DATA_BLOCK "DB_ALARM"   // DB100
{ S7_Optimized_Access := 'FALSE' }
// stored: AutoNumber false
   VAR
      ALARM : Struct
         ALARM_GLOBAL : Bool;   // globální alarm
         HERMA_ERROR : Bool;
         ALARM_2 : Bool;
         ALARM_3 : Bool;
         ALARM_4 : Bool;
         ALARM_5 : Bool;
         air : Bool;   // nedostatečný tlak vzduchu
         ALARM_7 : Bool;
         ALARM_8 : Bool;
         ALARM_9 : Bool;
         ALARM_10 : Bool;
         ALARM_11 : Bool;
         ALARM_12 : Bool;
         ALARM_13 : Bool;
         ALARM_14 : Bool;
         vypadek_safety_karty : Bool;
      END_STRUCT;
      WRONG : Struct
         NENI_INICIALIZACE : Bool;
         WRONG_global : Bool;
         dvere_L_tevreny : Bool;
         dvere_P_otevreny : Bool;
         WRONG_4 : Bool;
         WRONG_5 : Bool;
         WRONG_6 : Bool;
         WRONG_7 : Bool;
         WRONG_8 : Bool;
         WRONG_9 : Bool;
         WRONG_10 : Bool;
         WRONG_11 : Bool;
         WRONG_12 : Bool;
         WRONG_13 : Bool;
         rop_glob_warning : Bool;
         rop_active_autocale : Bool;
      END_STRUCT;
      OP0 : Struct
         ALARM : Struct
            DOOR_ERROR : Bool;
            ALARM_1 : Bool;
            ALARM_2 : Bool;
            ALARM_3 : Bool;
            ALARM_4 : Bool;
            ALARM_5 : Bool;
            ALARM_6 : Bool;
            ALARM_7 : Bool;
            ALARM_8 : Bool;
            ALARM_9 : Bool;
            ALARM_10 : Bool;
            ALARM_11 : Bool;
            ALARM_12 : Bool;
            ALARM_13 : Bool;
            ALARM_14 : Bool;
            ALARM_15 : Bool;
         END_STRUCT;
         WRONG : Struct
            WRONG_0 : Bool;
            WRONG_1 : Bool;
            WRONG_2 : Bool;
            WRONG_3 : Bool;
            WRONG_4 : Bool;
            WRONG_5 : Bool;
            WRONG_6 : Bool;
            WRONG_7 : Bool;
            WRONG_8 : Bool;
            WRONG_9 : Bool;
            WRONG_10 : Bool;
            WRONG_11 : Bool;
            WRONG_12 : Bool;
            WRONG_13 : Bool;
            WRONG_14 : Bool;
            WRONG_15 : Bool;
         END_STRUCT;
         M_0 : Int;
         M_1 : Int;
         M_2 : Int;
         M_3 : Int;
         M_4 : Int;
         M_5 : Int;
         M_6 : Int;
         M_7 : Int;
         M_8 : Int;
         M_9 : Int;
         M_10 : Int;
         M_11 : Int;
         M_12 : Int;
         M_13 : Int;
         M_14 : Int;
         M_15 : Int;
      END_STRUCT;
      OP1 : Struct
         ALARM : Struct
            dvere_1 : Bool;
            ALARM_1 : Bool;
            ALARM_2 : Bool;
            ALARM_3 : Bool;
            ALARM_4 : Bool;
            ALARM_5 : Bool;
            ALARM_6 : Bool;
            hladina_mimo_mez : Bool;
            ALARM_8 : Bool;
            ALARM_9 : Bool;
            ALARM_10 : Bool;
            ALARM_11 : Bool;
            ALARM_12 : Bool;
            ALARM_13 : Bool;
            ALARM_14 : Bool;
            ALARM_15 : Bool;
         END_STRUCT;
         WRONG : Struct
            WRONG_0 : Bool;
            WRONG_1 : Bool;
            WRONG_2 : Bool;
            WRONG_3 : Bool;
            WRONG_4 : Bool;
            WRONG_5 : Bool;
            WRONG_6 : Bool;
            WRONG_7 : Bool;
            WRONG_8 : Bool;
            WRONG_9 : Bool;
            WRONG_10 : Bool;
            WRONG_11 : Bool;
            WRONG_12 : Bool;
            WRONG_13 : Bool;
            WRONG_14 : Bool;
            WRONG_15 : Bool;
         END_STRUCT;
         "-Y7_KARUSEL" : Int;
         "-Y9_ZARAZKA" : Int;
         M_2 : Int;
         M_3 : Int;
         M_4 : Int;
         M_5 : Int;
         M_6 : Int;
         M_7 : Int;
         M_8 : Int;
         M_9 : Int;
         M_10 : Int;
         M_11 : Int;
         M_12 : Int;
         M_13 : Int;
         M_14 : Int;
         M_15 : Int;
      END_STRUCT;
      OP2 : Struct
         ALARM : Struct
            dvere_1 : Bool;
            dvere_2 : Bool;
            dvere_3 : Bool;
            dvere_4 : Bool;
            paprsek : Bool;
            porucha_svarovani : Bool;
            rop_alarm : Bool;
            servo_power_error : Bool;
            servo_jog_error : Bool;
            servo_homing : Bool;
            Cel_podel_porucha : Bool;
            vysoka_tuzka : Bool;
            ALARM_12 : Bool;
            ALARM_13 : Bool;
            folie : Bool;
            ALARM_15 : Bool;
         END_STRUCT;
         WRONG : Struct
            WRONG_0 : Bool;
            WRONG_1 : Bool;
            WRONG_2 : Bool;
            WRONG_3 : Bool;
            WRONG_4 : Bool;
            WRONG_5 : Bool;
            WRONG_6 : Bool;
            WRONG_7 : Bool;
            WRONG_8 : Bool;
            WRONG_9 : Bool;
            WRONG_10 : Bool;
            WRONG_11 : Bool;
            WRONG_12 : Bool;
            WRONG_13 : Bool;
            WRONG_14 : Bool;
            WRONG_15 : Bool;
         END_STRUCT;
         A1 : Int;   // -YA1
         A2 : Int;   // -YA2
         A3 : Int;   // -YA3
         A4 : Int;   // -YA4
         A5 : Int;   // -YA5
         A6 : Int;   // -YA6
         A7 : Int;   // -YA7
         A8 : Int;   // -YA8
         M_8 : Int;
         M_9 : Int;
         M_10 : Int;
         M_11 : Int;
         M_12 : Int;
         M_13 : Int;
         M_14 : Int;
         M_15 : Int;
      END_STRUCT;
      OP3 : Struct
         ALARM : Struct
            ALARM_0 : Bool;
            ALARM_1 : Bool;
            ALARM_2 : Bool;
            ALARM_3 : Bool;
            ALARM_4 : Bool;
            ALARM_5 : Bool;
            ALARM_6 : Bool;
            ALARM_7 : Bool;
            ALARM_8 : Bool;
            ALARM_9 : Bool;
            ALARM_10 : Bool;
            ALARM_11 : Bool;
            ALARM_12 : Bool;
            ALARM_13 : Bool;
            ALARM_14 : Bool;
            ALARM_15 : Bool;
         END_STRUCT;
         WRONG : Struct
            WRONG_0 : Bool;
            WRONG_1 : Bool;
            WRONG_2 : Bool;
            WRONG_3 : Bool;
            WRONG_4 : Bool;
            WRONG_5 : Bool;
            WRONG_6 : Bool;
            WRONG_7 : Bool;
            WRONG_8 : Bool;
            WRONG_9 : Bool;
            WRONG_10 : Bool;
            WRONG_11 : Bool;
            WRONG_12 : Bool;
            WRONG_13 : Bool;
            WRONG_14 : Bool;
            WRONG_15 : Bool;
         END_STRUCT;
         B1 : Int;   // -YB1
         B2 : Int;   // -YB2
         B3 : Int;   // -YB3
         B4 : Int;   // -YB4
         B5 : Int;   // -YB5
         B6 : Int;   // -YB6
         B7 : Int;   // -YB7
         B8 : Int;   // -YB8
         M_8 : Int;
         M_9 : Int;
         M_10 : Int;
         M_11 : Int;
         M_12 : Int;
         M_13 : Int;
         M_14 : Int;
         M_15 : Int;
      END_STRUCT;
      OP4 : Struct
         ALARM : Struct
            odsavani_nefunguje : Bool;
            ALARM_1 : Bool;
            ALARM_2 : Bool;
            ALARM_3 : Bool;
            ALARM_4 : Bool;
            ALARM_5 : Bool;
            ALARM_6 : Bool;
            ALARM_7 : Bool;
            ALARM_8 : Bool;
            ALARM_9 : Bool;
            ALARM_10 : Bool;
            ALARM_11 : Bool;
            ALARM_12 : Bool;
            ALARM_13 : Bool;
            ALARM_14 : Bool;
            ALARM_15 : Bool;
         END_STRUCT;
         WRONG : Struct
            WRONG_0 : Bool;
            WRONG_1 : Bool;
            WRONG_2 : Bool;
            WRONG_3 : Bool;
            WRONG_4 : Bool;
            WRONG_5 : Bool;
            WRONG_6 : Bool;
            WRONG_7 : Bool;
            WRONG_8 : Bool;
            WRONG_9 : Bool;
            WRONG_10 : Bool;
            WRONG_11 : Bool;
            WRONG_12 : Bool;
            WRONG_13 : Bool;
            WRONG_14 : Bool;
            WRONG_15 : Bool;
         END_STRUCT;
         M_0 : Int;
         M_1 : Int;
         M_2 : Int;
         M_3 : Int;
         M_4 : Int;
         M_5 : Int;
         M_6 : Int;
         M_7 : Int;
         M_8 : Int;
         M_9 : Int;
         M_10 : Int;
         M_11 : Int;
         M_12 : Int;
         M_13 : Int;
         M_14 : Int;
         M_15 : Int;
      END_STRUCT;
      OP5 : Struct
         ALARM : Struct
            ALARM_0 : Bool;
            ALARM_1 : Bool;
            ALARM_2 : Bool;
            ALARM_3 : Bool;
            ALARM_4 : Bool;
            ALARM_5 : Bool;
            ALARM_6 : Bool;
            ALARM_7 : Bool;
            ALARM_8 : Bool;
            ALARM_9 : Bool;
            ALARM_10 : Bool;
            ALARM_11 : Bool;
            ALARM_12 : Bool;
            ALARM_13 : Bool;
            ALARM_14 : Bool;
            ALARM_15 : Bool;
         END_STRUCT;
         WRONG : Struct
            WRONG_0 : Bool;
            WRONG_1 : Bool;
            WRONG_2 : Bool;
            WRONG_3 : Bool;
            WRONG_4 : Bool;
            WRONG_5 : Bool;
            WRONG_6 : Bool;
            WRONG_7 : Bool;
            WRONG_8 : Bool;
            WRONG_9 : Bool;
            WRONG_10 : Bool;
            WRONG_11 : Bool;
            WRONG_12 : Bool;
            WRONG_13 : Bool;
            WRONG_14 : Bool;
            WRONG_15 : Bool;
         END_STRUCT;
         M_0 : Int;
         M_1 : Int;
         M_2 : Int;
         M_3 : Int;
         M_4 : Int;
         M_5 : Int;
         M_6 : Int;
         M_7 : Int;
         M_8 : Int;
         M_9 : Int;
         M_10 : Int;
         M_11 : Int;
         M_12 : Int;
         M_13 : Int;
         M_14 : Int;
         M_15 : Int;
      END_STRUCT;
      null : Struct
         ALARM_0 : Bool;
         ALARM_1 : Bool;
         ALARM_2 : Bool;
         ALARM_3 : Bool;
         ALARM_4 : Bool;
         ALARM_5 : Bool;
         ALARM_6 : Bool;
         ALARM_7 : Bool;
         ALARM_8 : Bool;
         ALARM_9 : Bool;
         ALARM_10 : Bool;
         ALARM_11 : Bool;
         ALARM_12 : Bool;
         ALARM_13 : Bool;
         ALARM_14 : Bool;
         ALARM_15 : Bool;
      END_STRUCT;
      alarmy : Array[0..255] of Bool;
      alarm_line : Int;
      wrong_line : Int;
      alarm_op_1 : Int;
      wrong_op_1 : Int;
      alarm_op_2 : Int;
      wrong_op_2 : Int;
      alarm_op_3 : Int;
      wrong_op_3 : Int;
      alarm_op_4 : Int;
      wrong_op_4 : Int;
      alarm_op_5 : Int;
      wrong_op_5 : Int;
      T_tiskarna : TON_TIME;
   END_VAR
BEGIN
END_DATA_BLOCK

DATA_BLOCK "DB_STS_M"   // DB101
{ S7_Optimized_Access := 'FALSE' }
// stored: AutoNumber false
   VAR
      OP0 : Struct
         STS_M0 : UInt;
         STS_M1 : UInt;
         STS_M2 : UInt;
         STS_M3 : UInt;
         STS_M4 : UInt;
         STS_M5 : UInt;
         STS_M6 : UInt;
         STS_M7 : UInt;
         STS_M8 : UInt;
         STS_M9 : UInt;
         STS_M10 : UInt;
         STS_M11 : UInt;
         STS_M12 : UInt;
         STS_M13 : UInt;
         STS_M14 : UInt;
         STS_M15 : UInt;
      END_STRUCT;
      OP1 : Struct
         KARUSEL : UInt;
         ZARAZKA : UInt;
         STS_M2 : UInt;
         STS_M3 : UInt;
         STS_M4 : UInt;
         STS_M5 : UInt;
         STS_M6 : UInt;
         STS_M7 : UInt;
         STS_M8 : UInt;
         STS_M9 : UInt;
         STS_M10 : UInt;
         STS_M11 : UInt;
         STS_M12 : UInt;
         STS_M13 : UInt;
         STS_M14 : UInt;
         STS_M15 : UInt;
         OP1 : Struct
            STS_M0 : UInt;
            STS_M1 : UInt;
            STS_M2 : UInt;
            STS_M3 : UInt;
            STS_M4 : UInt;
            STS_M5 : UInt;
            STS_M6 : UInt;
            STS_M7 : UInt;
            STS_M8 : UInt;
            STS_M9 : UInt;
            STS_M10 : UInt;
            STS_M11 : UInt;
            STS_M12 : UInt;
            STS_M13 : UInt;
            STS_M14 : UInt;
            STS_M15 : UInt;
         END_STRUCT;
      END_STRUCT;
      OP2 : Struct
         A1 : UInt;
         A2 : UInt;
         A3 : UInt;
         A4 : UInt;
         A5 : UInt;
         A6 : UInt;
         A7 : UInt;
         A8 : UInt;
         STS_M8 : UInt;
         STS_M9 : UInt;
         STS_M10 : UInt;
         STS_M11 : UInt;
         STS_M12 : UInt;
         STS_M13 : UInt;
         STS_M14 : UInt;
         STS_M15 : UInt;
      END_STRUCT;
      OP3 : Struct
         B1 : UInt;
         B2 : UInt;
         B3 : UInt;
         B4 : UInt;
         B5 : UInt;
         B6 : UInt;
         B7 : UInt;
         B8 : UInt;
         STS_M8 : UInt;
         STS_M9 : UInt;
         STS_M10 : UInt;
         STS_M11 : UInt;
         STS_M12 : UInt;
         STS_M13 : UInt;
         STS_M14 : UInt;
         STS_M15 : UInt;
      END_STRUCT;
   END_VAR
BEGIN
END_DATA_BLOCK

DATA_BLOCK "DB_DATA_LASER"   // DB401
{ S7_Optimized_Access := 'TRUE' }
// stored: AutoNumber false, MemoryReserve 100
   VAR
      LASER_DATA_READ : Array[0..71] of Byte;
      LASER_DATA_WRITE : Array[0..71] of Byte;
      READ : Bool;
      WRITE : Bool;
   END_VAR
BEGIN
END_DATA_BLOCK

DATA_BLOCK "DB_LASER"   // DB402
{ S7_Optimized_Access := 'TRUE' }
// stored: AutoNumber false, MemoryReserve 100
   VAR
      DATA_DO_ETIKETY : Struct
         TEXT : String[5];
         "INT" : Int;
         "REAL" : Real;
         PROGRAM : Array[0..1] of String[10];
      END_STRUCT;
      DATA_DO_DAT : Struct
         ZAVORKA_L : Char := '<';
         ZAVORKA_P : Char := '>';
         XLP : Array[0..3] of Char;
      END_STRUCT;
      smaz_me_start : Bool;
      smaz_me_adresa : Int;
   END_VAR
BEGIN
   DATA_DO_ETIKETY.PROGRAM[0] := 'TEST_1';
   DATA_DO_ETIKETY.PROGRAM[1] := 'TEST_222';
   DATA_DO_DAT.XLP[0] := '.';
   DATA_DO_DAT.XLP[1] := 'x';
   DATA_DO_DAT.XLP[2] := 'l';
   DATA_DO_DAT.XLP[3] := 'p';
END_DATA_BLOCK

ORGANIZATION_BLOCK "Main"   // OB1, LAD, ProgramCycle
TITLE = "Main Program Sweep (Cycle)"
{ S7_Optimized_Access := 'TRUE' }
// stored: SetENOAutomatically false
   VAR_INPUT
      Initial_Call : Bool;   // Initial call of this OB
      Remanence : Bool;   // =True, if remanent data are available
   END_VAR
BEGIN

REGION Network 1
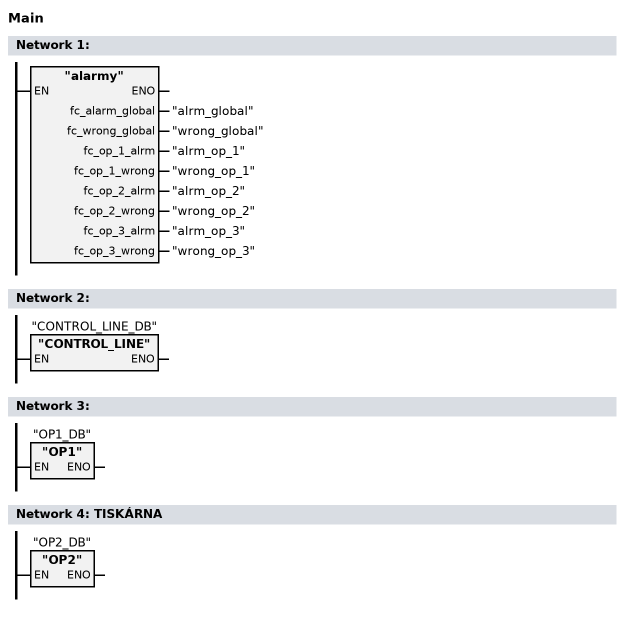
   RUNG wire#powerrail
      "alarmy"(fc_alarm_global => "alrm_global", fc_wrong_global => "wrong_global", fc_op_1_alrm => "alrm_op_1", fc_op_1_wrong => "wrong_op_1", fc_op_2_alrm => "alrm_op_2", fc_op_2_wrong => "wrong_op_2", fc_op_3_alrm => "alrm_op_3", fc_op_3_wrong => "wrong_op_3")
   END_RUNG
   // the same network as SCL:
   "alarmy"(fc_alarm_global => "alrm_global",
            fc_wrong_global => "wrong_global",
            fc_op_1_alrm => "alrm_op_1",
            fc_op_1_wrong => "wrong_op_1",
            fc_op_2_alrm => "alrm_op_2",
            fc_op_2_wrong => "wrong_op_2",
            fc_op_3_alrm => "alrm_op_3",
            fc_op_3_wrong => "wrong_op_3");
END_REGION

REGION Network 2
   RUNG wire#powerrail
      "CONTROL_LINE_DB"()
   END_RUNG
   // the same network as SCL:
   "CONTROL_LINE_DB"();   // "CONTROL_LINE"
END_REGION

REGION Network 3
   RUNG wire#powerrail
      "OP1_DB"()
   END_RUNG
   // the same network as SCL:
   "OP1_DB"();   // "OP1"
END_REGION

REGION Network 4: TISKÁRNA
   RUNG wire#powerrail
      "OP2_DB"()
   END_RUNG
   // the same network as SCL:
   "OP2_DB"();   // "OP2"
END_REGION
END_ORGANIZATION_BLOCK

FUNCTION "alarmy" : Void   // FC100, LAD
{ S7_Optimized_Access := 'TRUE' }
// stored: AutoNumber false, SetENOAutomatically false
   VAR_OUTPUT
      fc_alarm_global : Bool;
      fc_wrong_global : Bool;
      fc_op_1_alrm : Bool;
      fc_op_1_wrong : Bool;
      fc_op_2_alrm : Bool;
      fc_op_2_wrong : Bool;
      fc_op_3_alrm : Bool;
      fc_op_3_wrong : Bool;
   END_VAR
   VAR_TEMP
      OP_1_E : Bool;
      OP_2_E : Bool;
      OP_3_E : Bool;
      OP_4_E : Bool;
      OP_5_E : Bool;
      OP_1_W : Bool;
      OP_2_W : Bool;
      OP_3_W : Bool;
      OP_4_W : Bool;
      OP_5_W : Bool;
   END_VAR
   VAR CONSTANT
      TIME_ERROR_BOR : Time := T#4S;
   END_VAR
BEGIN

REGION Network 1: op_1 alarmy proces
END_REGION

REGION Network 2: op_1_warning_proces
END_REGION

REGION Network 3: OP_1_ALARM
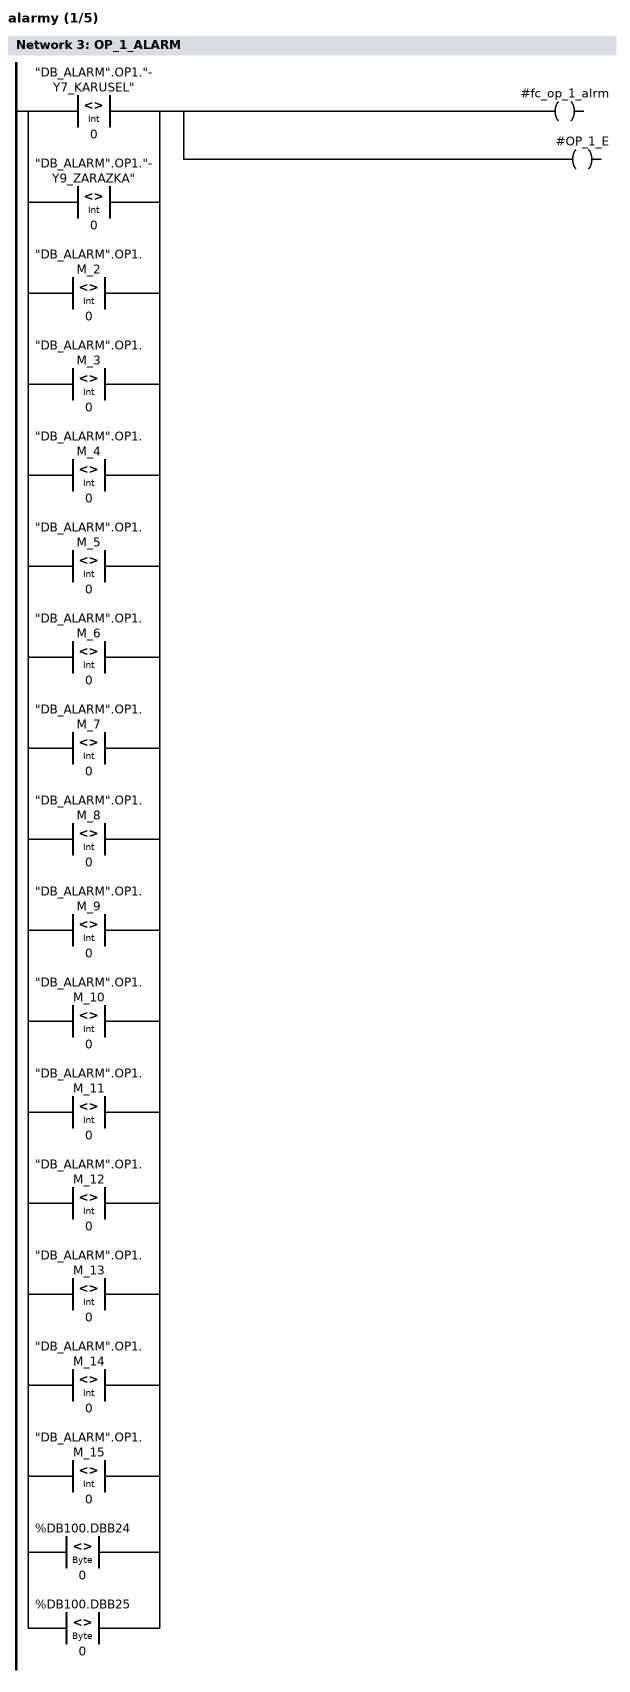
   RUNG wire#powerrail
      { S7_Templates := "SrcType := Int" } NE_Contact(in1 := "DB_ALARM".OP1."-Y7_KARUSEL", in2 := 0)
      wire#w1
      Coil( #fc_op_1_alrm )
   END_RUNG
   RUNG wire#powerrail
      { S7_Templates := "SrcType := Int" } NE_Contact(in1 := "DB_ALARM".OP1."-Y9_ZARAZKA", in2 := 0)
   END_RUNG wire#w1
   RUNG wire#powerrail
      { S7_Templates := "SrcType := Int" } NE_Contact(in1 := "DB_ALARM".OP1.M_2, in2 := 0)
   END_RUNG wire#w1
   RUNG wire#powerrail
      { S7_Templates := "SrcType := Int" } NE_Contact(in1 := "DB_ALARM".OP1.M_3, in2 := 0)
   END_RUNG wire#w1
   RUNG wire#powerrail
      { S7_Templates := "SrcType := Int" } NE_Contact(in1 := "DB_ALARM".OP1.M_4, in2 := 0)
   END_RUNG wire#w1
   RUNG wire#powerrail
      { S7_Templates := "SrcType := Int" } NE_Contact(in1 := "DB_ALARM".OP1.M_5, in2 := 0)
   END_RUNG wire#w1
   RUNG wire#powerrail
      { S7_Templates := "SrcType := Int" } NE_Contact(in1 := "DB_ALARM".OP1.M_6, in2 := 0)
   END_RUNG wire#w1
   RUNG wire#powerrail
      { S7_Templates := "SrcType := Int" } NE_Contact(in1 := "DB_ALARM".OP1.M_7, in2 := 0)
   END_RUNG wire#w1
   RUNG wire#powerrail
      { S7_Templates := "SrcType := Int" } NE_Contact(in1 := "DB_ALARM".OP1.M_8, in2 := 0)
   END_RUNG wire#w1
   RUNG wire#powerrail
      { S7_Templates := "SrcType := Int" } NE_Contact(in1 := "DB_ALARM".OP1.M_9, in2 := 0)
   END_RUNG wire#w1
   RUNG wire#powerrail
      { S7_Templates := "SrcType := Int" } NE_Contact(in1 := "DB_ALARM".OP1.M_10, in2 := 0)
   END_RUNG wire#w1
   RUNG wire#powerrail
      { S7_Templates := "SrcType := Int" } NE_Contact(in1 := "DB_ALARM".OP1.M_11, in2 := 0)
   END_RUNG wire#w1
   RUNG wire#powerrail
      { S7_Templates := "SrcType := Int" } NE_Contact(in1 := "DB_ALARM".OP1.M_12, in2 := 0)
   END_RUNG wire#w1
   RUNG wire#powerrail
      { S7_Templates := "SrcType := Int" } NE_Contact(in1 := "DB_ALARM".OP1.M_13, in2 := 0)
   END_RUNG wire#w1
   RUNG wire#powerrail
      { S7_Templates := "SrcType := Int" } NE_Contact(in1 := "DB_ALARM".OP1.M_14, in2 := 0)
   END_RUNG wire#w1
   RUNG wire#powerrail
      { S7_Templates := "SrcType := Int" } NE_Contact(in1 := "DB_ALARM".OP1.M_15, in2 := 0)
   END_RUNG wire#w1
   RUNG wire#powerrail
      { S7_Templates := "SrcType := Byte" } NE_Contact(in1 := %DB100.DBB24, in2 := 0)
   END_RUNG wire#w1
   RUNG wire#powerrail
      { S7_Templates := "SrcType := Byte" } NE_Contact(in1 := %DB100.DBB25, in2 := 0)
   END_RUNG wire#w1
   RUNG wire#w1
      Coil( #OP_1_E )
   END_RUNG
   // the same network as SCL:
   #fc_op_1_alrm := ("DB_ALARM".OP1."-Y7_KARUSEL" <> 0) OR ("DB_ALARM".OP1."-Y9_ZARAZKA" <> 0) OR ("DB_ALARM".OP1.M_2 <> 0) OR ("DB_ALARM".OP1.M_3 <> 0) OR ("DB_ALARM".OP1.M_4 <> 0) OR ("DB_ALARM".OP1.M_5 <> 0) OR ("DB_ALARM".OP1.M_6 <> 0) OR ("DB_ALARM".OP1.M_7 <> 0) OR ("DB_ALARM".OP1.M_8 <> 0) OR ("DB_ALARM".OP1.M_9 <> 0) OR ("DB_ALARM".OP1.M_10 <> 0) OR ("DB_ALARM".OP1.M_11 <> 0) OR ("DB_ALARM".OP1.M_12 <> 0) OR ("DB_ALARM".OP1.M_13 <> 0) OR ("DB_ALARM".OP1.M_14 <> 0) OR ("DB_ALARM".OP1.M_15 <> 0) OR (%DB100.DBB24 <> 0) OR (%DB100.DBB25 <> 0);
   #OP_1_E := #fc_op_1_alrm;
END_REGION

REGION Network 4: OP_2_ALARM
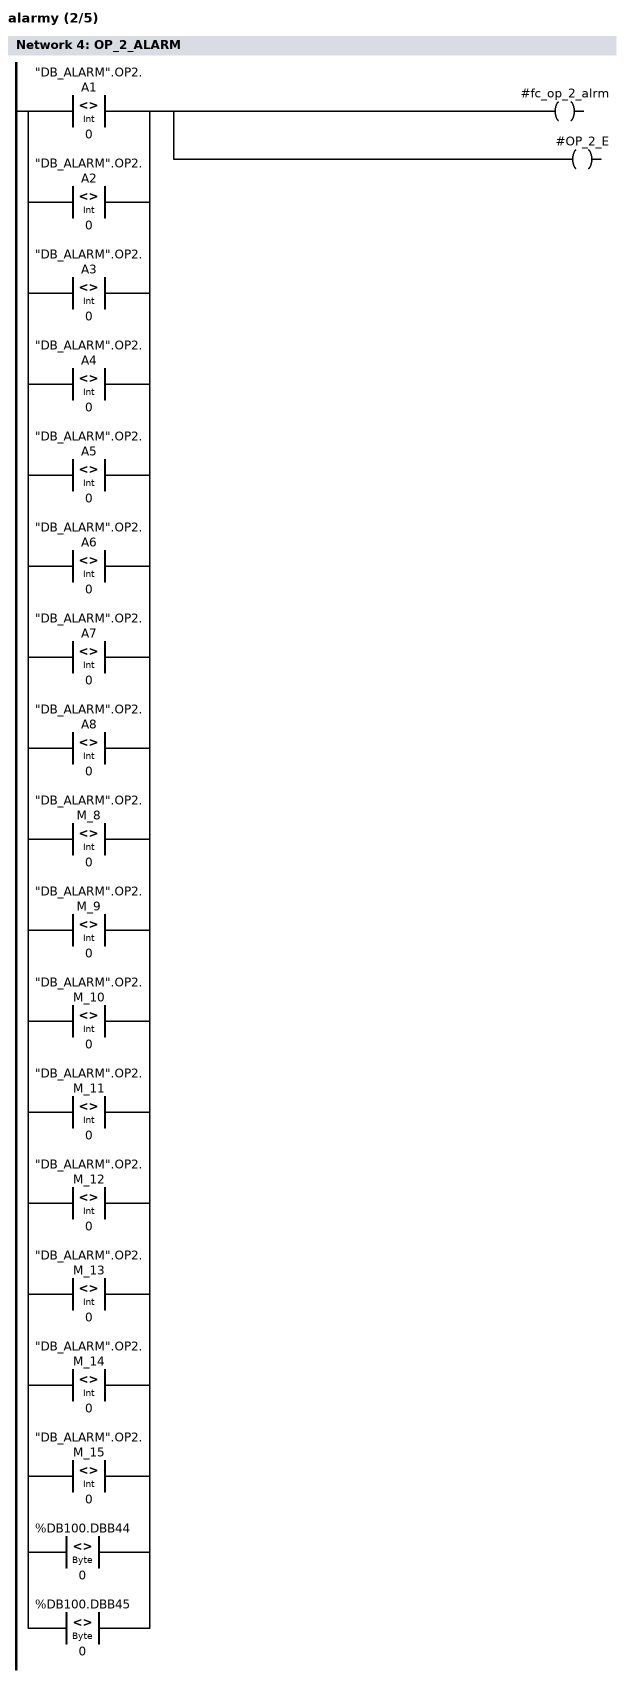
   RUNG wire#powerrail
      { S7_Templates := "SrcType := Int" } NE_Contact(in1 := "DB_ALARM".OP2.A1, in2 := 0)
      wire#w1
      Coil( #fc_op_2_alrm )
   END_RUNG
   RUNG wire#powerrail
      { S7_Templates := "SrcType := Int" } NE_Contact(in1 := "DB_ALARM".OP2.A2, in2 := 0)
   END_RUNG wire#w1
   RUNG wire#powerrail
      { S7_Templates := "SrcType := Int" } NE_Contact(in1 := "DB_ALARM".OP2.A3, in2 := 0)
   END_RUNG wire#w1
   RUNG wire#powerrail
      { S7_Templates := "SrcType := Int" } NE_Contact(in1 := "DB_ALARM".OP2.A4, in2 := 0)
   END_RUNG wire#w1
   RUNG wire#powerrail
      { S7_Templates := "SrcType := Int" } NE_Contact(in1 := "DB_ALARM".OP2.A5, in2 := 0)
   END_RUNG wire#w1
   RUNG wire#powerrail
      { S7_Templates := "SrcType := Int" } NE_Contact(in1 := "DB_ALARM".OP2.A6, in2 := 0)
   END_RUNG wire#w1
   RUNG wire#powerrail
      { S7_Templates := "SrcType := Int" } NE_Contact(in1 := "DB_ALARM".OP2.A7, in2 := 0)
   END_RUNG wire#w1
   RUNG wire#powerrail
      { S7_Templates := "SrcType := Int" } NE_Contact(in1 := "DB_ALARM".OP2.A8, in2 := 0)
   END_RUNG wire#w1
   RUNG wire#powerrail
      { S7_Templates := "SrcType := Int" } NE_Contact(in1 := "DB_ALARM".OP2.M_8, in2 := 0)
   END_RUNG wire#w1
   RUNG wire#powerrail
      { S7_Templates := "SrcType := Int" } NE_Contact(in1 := "DB_ALARM".OP2.M_9, in2 := 0)
   END_RUNG wire#w1
   RUNG wire#powerrail
      { S7_Templates := "SrcType := Int" } NE_Contact(in1 := "DB_ALARM".OP2.M_10, in2 := 0)
   END_RUNG wire#w1
   RUNG wire#powerrail
      { S7_Templates := "SrcType := Int" } NE_Contact(in1 := "DB_ALARM".OP2.M_11, in2 := 0)
   END_RUNG wire#w1
   RUNG wire#powerrail
      { S7_Templates := "SrcType := Int" } NE_Contact(in1 := "DB_ALARM".OP2.M_12, in2 := 0)
   END_RUNG wire#w1
   RUNG wire#powerrail
      { S7_Templates := "SrcType := Int" } NE_Contact(in1 := "DB_ALARM".OP2.M_13, in2 := 0)
   END_RUNG wire#w1
   RUNG wire#powerrail
      { S7_Templates := "SrcType := Int" } NE_Contact(in1 := "DB_ALARM".OP2.M_14, in2 := 0)
   END_RUNG wire#w1
   RUNG wire#powerrail
      { S7_Templates := "SrcType := Int" } NE_Contact(in1 := "DB_ALARM".OP2.M_15, in2 := 0)
   END_RUNG wire#w1
   RUNG wire#powerrail
      { S7_Templates := "SrcType := Byte" } NE_Contact(in1 := %DB100.DBB44, in2 := 0)
   END_RUNG wire#w1
   RUNG wire#powerrail
      { S7_Templates := "SrcType := Byte" } NE_Contact(in1 := %DB100.DBB45, in2 := 0)
   END_RUNG wire#w1
   RUNG wire#w1
      Coil( #OP_2_E )
   END_RUNG
   // the same network as SCL:
   #fc_op_2_alrm := ("DB_ALARM".OP2.A1 <> 0) OR ("DB_ALARM".OP2.A2 <> 0) OR ("DB_ALARM".OP2.A3 <> 0) OR ("DB_ALARM".OP2.A4 <> 0) OR ("DB_ALARM".OP2.A5 <> 0) OR ("DB_ALARM".OP2.A6 <> 0) OR ("DB_ALARM".OP2.A7 <> 0) OR ("DB_ALARM".OP2.A8 <> 0) OR ("DB_ALARM".OP2.M_8 <> 0) OR ("DB_ALARM".OP2.M_9 <> 0) OR ("DB_ALARM".OP2.M_10 <> 0) OR ("DB_ALARM".OP2.M_11 <> 0) OR ("DB_ALARM".OP2.M_12 <> 0) OR ("DB_ALARM".OP2.M_13 <> 0) OR ("DB_ALARM".OP2.M_14 <> 0) OR ("DB_ALARM".OP2.M_15 <> 0) OR (%DB100.DBB44 <> 0) OR (%DB100.DBB45 <> 0);
   #OP_2_E := #fc_op_2_alrm;
END_REGION

REGION Network 5: OP_3_ALARM
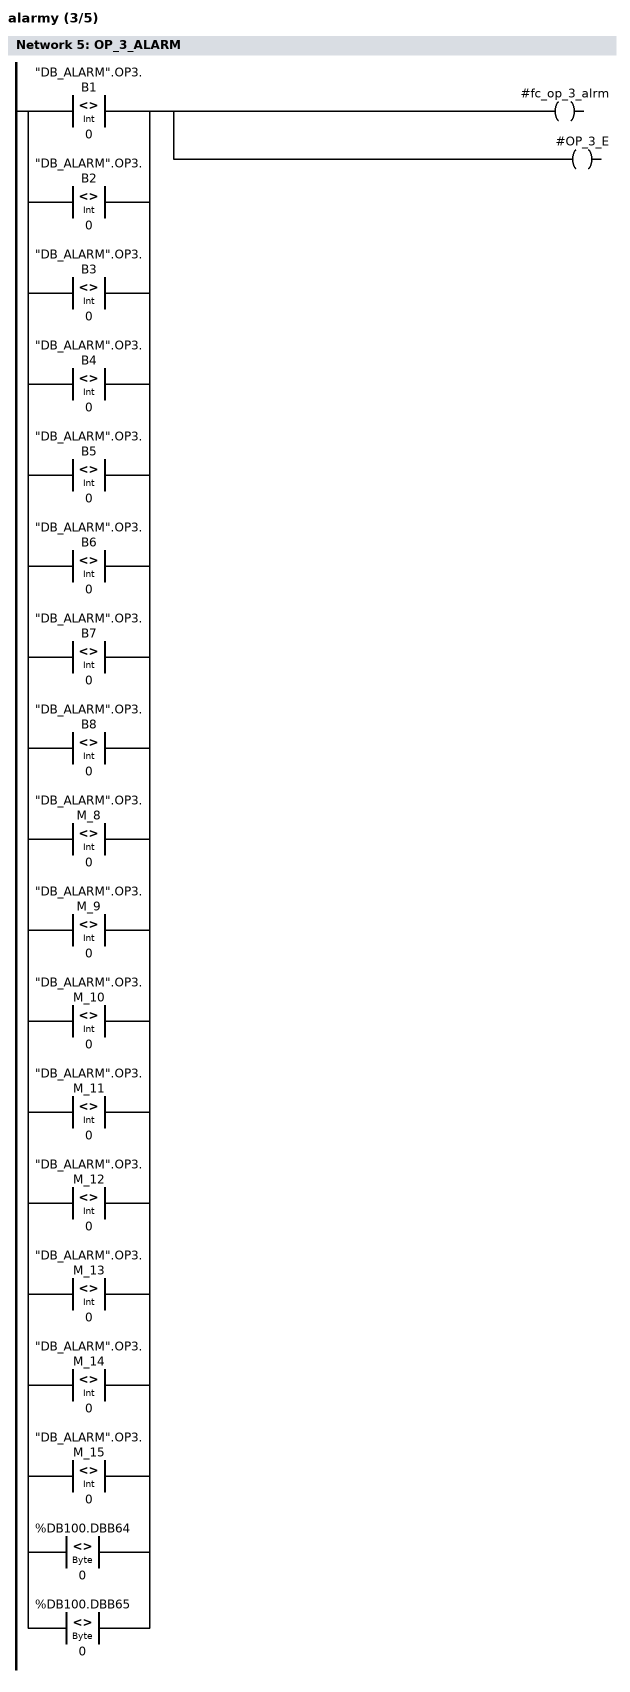
   RUNG wire#powerrail
      { S7_Templates := "SrcType := Int" } NE_Contact(in1 := "DB_ALARM".OP3.B1, in2 := 0)
      wire#w1
      Coil( #fc_op_3_alrm )
   END_RUNG
   RUNG wire#powerrail
      { S7_Templates := "SrcType := Int" } NE_Contact(in1 := "DB_ALARM".OP3.B2, in2 := 0)
   END_RUNG wire#w1
   RUNG wire#powerrail
      { S7_Templates := "SrcType := Int" } NE_Contact(in1 := "DB_ALARM".OP3.B3, in2 := 0)
   END_RUNG wire#w1
   RUNG wire#powerrail
      { S7_Templates := "SrcType := Int" } NE_Contact(in1 := "DB_ALARM".OP3.B4, in2 := 0)
   END_RUNG wire#w1
   RUNG wire#powerrail
      { S7_Templates := "SrcType := Int" } NE_Contact(in1 := "DB_ALARM".OP3.B5, in2 := 0)
   END_RUNG wire#w1
   RUNG wire#powerrail
      { S7_Templates := "SrcType := Int" } NE_Contact(in1 := "DB_ALARM".OP3.B6, in2 := 0)
   END_RUNG wire#w1
   RUNG wire#powerrail
      { S7_Templates := "SrcType := Int" } NE_Contact(in1 := "DB_ALARM".OP3.B7, in2 := 0)
   END_RUNG wire#w1
   RUNG wire#powerrail
      { S7_Templates := "SrcType := Int" } NE_Contact(in1 := "DB_ALARM".OP3.B8, in2 := 0)
   END_RUNG wire#w1
   RUNG wire#powerrail
      { S7_Templates := "SrcType := Int" } NE_Contact(in1 := "DB_ALARM".OP3.M_8, in2 := 0)
   END_RUNG wire#w1
   RUNG wire#powerrail
      { S7_Templates := "SrcType := Int" } NE_Contact(in1 := "DB_ALARM".OP3.M_9, in2 := 0)
   END_RUNG wire#w1
   RUNG wire#powerrail
      { S7_Templates := "SrcType := Int" } NE_Contact(in1 := "DB_ALARM".OP3.M_10, in2 := 0)
   END_RUNG wire#w1
   RUNG wire#powerrail
      { S7_Templates := "SrcType := Int" } NE_Contact(in1 := "DB_ALARM".OP3.M_11, in2 := 0)
   END_RUNG wire#w1
   RUNG wire#powerrail
      { S7_Templates := "SrcType := Int" } NE_Contact(in1 := "DB_ALARM".OP3.M_12, in2 := 0)
   END_RUNG wire#w1
   RUNG wire#powerrail
      { S7_Templates := "SrcType := Int" } NE_Contact(in1 := "DB_ALARM".OP3.M_13, in2 := 0)
   END_RUNG wire#w1
   RUNG wire#powerrail
      { S7_Templates := "SrcType := Int" } NE_Contact(in1 := "DB_ALARM".OP3.M_14, in2 := 0)
   END_RUNG wire#w1
   RUNG wire#powerrail
      { S7_Templates := "SrcType := Int" } NE_Contact(in1 := "DB_ALARM".OP3.M_15, in2 := 0)
   END_RUNG wire#w1
   RUNG wire#powerrail
      { S7_Templates := "SrcType := Byte" } NE_Contact(in1 := %DB100.DBB64, in2 := 0)
   END_RUNG wire#w1
   RUNG wire#powerrail
      { S7_Templates := "SrcType := Byte" } NE_Contact(in1 := %DB100.DBB65, in2 := 0)
   END_RUNG wire#w1
   RUNG wire#w1
      Coil( #OP_3_E )
   END_RUNG
   // the same network as SCL:
   #fc_op_3_alrm := ("DB_ALARM".OP3.B1 <> 0) OR ("DB_ALARM".OP3.B2 <> 0) OR ("DB_ALARM".OP3.B3 <> 0) OR ("DB_ALARM".OP3.B4 <> 0) OR ("DB_ALARM".OP3.B5 <> 0) OR ("DB_ALARM".OP3.B6 <> 0) OR ("DB_ALARM".OP3.B7 <> 0) OR ("DB_ALARM".OP3.B8 <> 0) OR ("DB_ALARM".OP3.M_8 <> 0) OR ("DB_ALARM".OP3.M_9 <> 0) OR ("DB_ALARM".OP3.M_10 <> 0) OR ("DB_ALARM".OP3.M_11 <> 0) OR ("DB_ALARM".OP3.M_12 <> 0) OR ("DB_ALARM".OP3.M_13 <> 0) OR ("DB_ALARM".OP3.M_14 <> 0) OR ("DB_ALARM".OP3.M_15 <> 0) OR (%DB100.DBB64 <> 0) OR (%DB100.DBB65 <> 0);
   #OP_3_E := #fc_op_3_alrm;
END_REGION

REGION Network 6: OP_1_WRONG
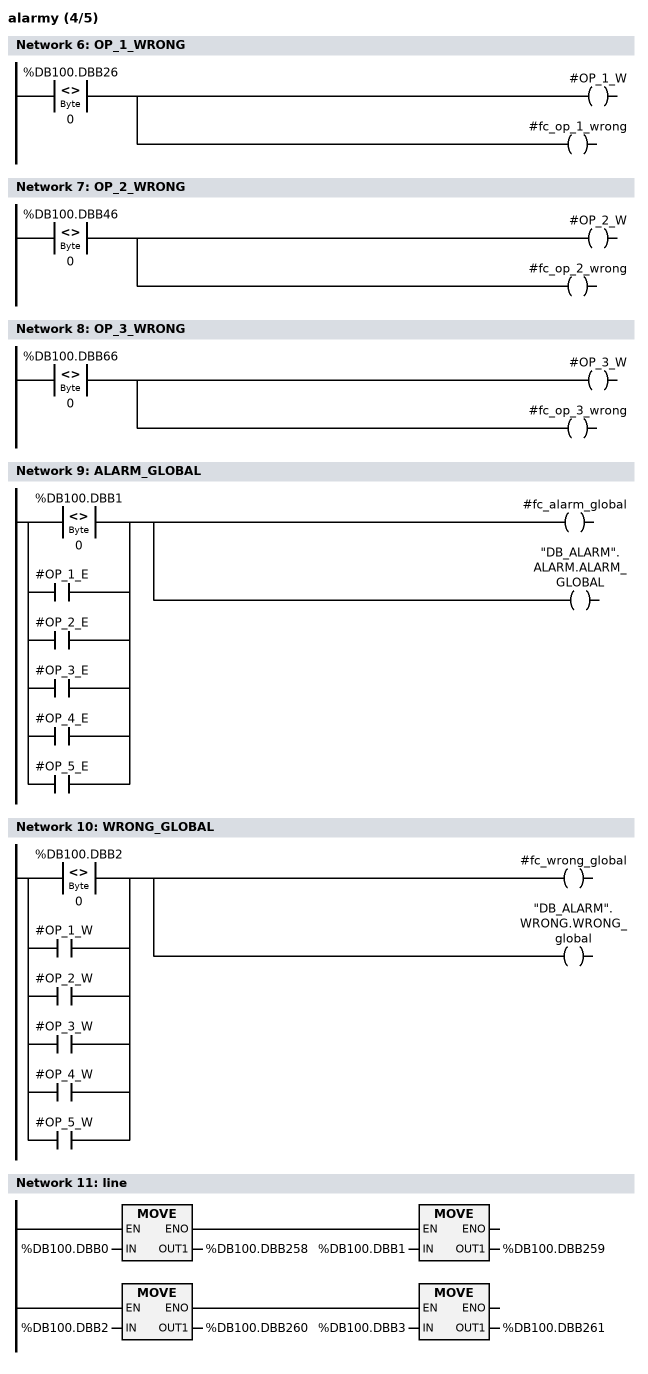
   RUNG wire#powerrail
      { S7_Templates := "SrcType := Byte" } NE_Contact(in1 := %DB100.DBB26, in2 := 0)
      wire#w1
      Coil( #OP_1_W )
   END_RUNG
   RUNG wire#w1
      Coil( #fc_op_1_wrong )
   END_RUNG
   // the same network as SCL:
   #OP_1_W := %DB100.DBB26 <> 0;
   #fc_op_1_wrong := #OP_1_W;
END_REGION

REGION Network 7: OP_2_WRONG
   RUNG wire#powerrail
      { S7_Templates := "SrcType := Byte" } NE_Contact(in1 := %DB100.DBB46, in2 := 0)
      wire#w1
      Coil( #OP_2_W )
   END_RUNG
   RUNG wire#w1
      Coil( #fc_op_2_wrong )
   END_RUNG
   // the same network as SCL:
   #OP_2_W := %DB100.DBB46 <> 0;
   #fc_op_2_wrong := #OP_2_W;
END_REGION

REGION Network 8: OP_3_WRONG
   RUNG wire#powerrail
      { S7_Templates := "SrcType := Byte" } NE_Contact(in1 := %DB100.DBB66, in2 := 0)
      wire#w1
      Coil( #OP_3_W )
   END_RUNG
   RUNG wire#w1
      Coil( #fc_op_3_wrong )
   END_RUNG
   // the same network as SCL:
   #OP_3_W := %DB100.DBB66 <> 0;
   #fc_op_3_wrong := #OP_3_W;
END_REGION

REGION Network 9: ALARM_GLOBAL
   RUNG wire#powerrail
      { S7_Templates := "SrcType := Byte" } NE_Contact(in1 := %DB100.DBB1, in2 := 0)
      wire#w1
      Coil( #fc_alarm_global )
   END_RUNG
   RUNG wire#powerrail
      Contact( #OP_1_E )
   END_RUNG wire#w1
   RUNG wire#powerrail
      Contact( #OP_2_E )
   END_RUNG wire#w1
   RUNG wire#powerrail
      Contact( #OP_3_E )
   END_RUNG wire#w1
   RUNG wire#powerrail
      Contact( #OP_4_E )
   END_RUNG wire#w1
   RUNG wire#powerrail
      Contact( #OP_5_E )
   END_RUNG wire#w1
   RUNG wire#w1
      Coil( "DB_ALARM".ALARM.ALARM_GLOBAL )
   END_RUNG
   // the same network as SCL:
   #fc_alarm_global := (%DB100.DBB1 <> 0) OR #OP_1_E OR #OP_2_E OR #OP_3_E OR #OP_4_E OR #OP_5_E;
   "DB_ALARM".ALARM.ALARM_GLOBAL := #fc_alarm_global;
END_REGION

REGION Network 10: WRONG_GLOBAL
   RUNG wire#powerrail
      { S7_Templates := "SrcType := Byte" } NE_Contact(in1 := %DB100.DBB2, in2 := 0)
      wire#w1
      Coil( #fc_wrong_global )
   END_RUNG
   RUNG wire#powerrail
      Contact( #OP_1_W )
   END_RUNG wire#w1
   RUNG wire#powerrail
      Contact( #OP_2_W )
   END_RUNG wire#w1
   RUNG wire#powerrail
      Contact( #OP_3_W )
   END_RUNG wire#w1
   RUNG wire#powerrail
      Contact( #OP_4_W )
   END_RUNG wire#w1
   RUNG wire#powerrail
      Contact( #OP_5_W )
   END_RUNG wire#w1
   RUNG wire#w1
      Coil( "DB_ALARM".WRONG.WRONG_global )
   END_RUNG
   // the same network as SCL:
   #fc_wrong_global := (%DB100.DBB2 <> 0) OR #OP_1_W OR #OP_2_W OR #OP_3_W OR #OP_4_W OR #OP_5_W;
   "DB_ALARM".WRONG.WRONG_global := #fc_wrong_global;
END_REGION

REGION Network 11: line
   RUNG wire#powerrail
      Move(in := %DB100.DBB0, out1 => %DB100.DBB258)
      Move(in := %DB100.DBB1, out1 => %DB100.DBB259)
   END_RUNG
   RUNG wire#powerrail
      Move(in := %DB100.DBB2, out1 => %DB100.DBB260)
      Move(in := %DB100.DBB3, out1 => %DB100.DBB261)
   END_RUNG
   // the same network as SCL:
   %DB100.DBB258 := %DB100.DBB0;
   %DB100.DBB259 := %DB100.DBB1;
   %DB100.DBB260 := %DB100.DBB2;
   %DB100.DBB261 := %DB100.DBB3;
END_REGION

REGION Network 12: op_1
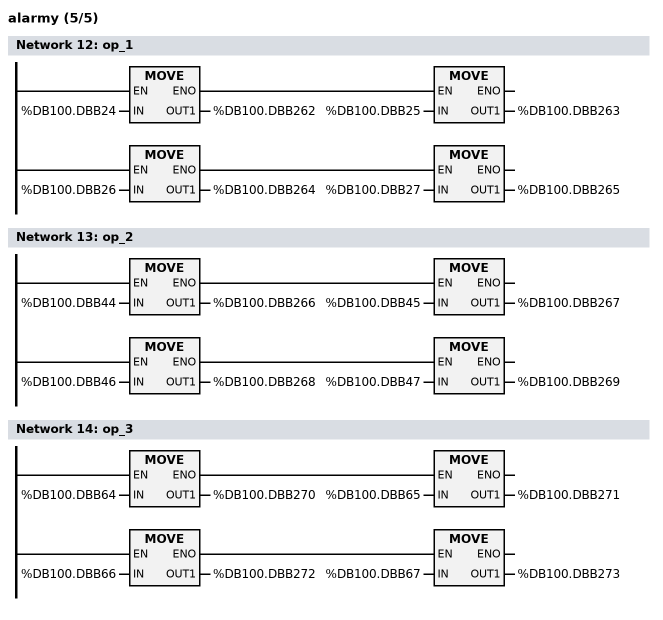
   RUNG wire#powerrail
      Move(in := %DB100.DBB24, out1 => %DB100.DBB262)
      Move(in := %DB100.DBB25, out1 => %DB100.DBB263)
   END_RUNG
   RUNG wire#powerrail
      Move(in := %DB100.DBB26, out1 => %DB100.DBB264)
      Move(in := %DB100.DBB27, out1 => %DB100.DBB265)
   END_RUNG
   // the same network as SCL:
   %DB100.DBB262 := %DB100.DBB24;
   %DB100.DBB263 := %DB100.DBB25;
   %DB100.DBB264 := %DB100.DBB26;
   %DB100.DBB265 := %DB100.DBB27;
END_REGION

REGION Network 13: op_2
   RUNG wire#powerrail
      Move(in := %DB100.DBB44, out1 => %DB100.DBB266)
      Move(in := %DB100.DBB45, out1 => %DB100.DBB267)
   END_RUNG
   RUNG wire#powerrail
      Move(in := %DB100.DBB46, out1 => %DB100.DBB268)
      Move(in := %DB100.DBB47, out1 => %DB100.DBB269)
   END_RUNG
   // the same network as SCL:
   %DB100.DBB266 := %DB100.DBB44;
   %DB100.DBB267 := %DB100.DBB45;
   %DB100.DBB268 := %DB100.DBB46;
   %DB100.DBB269 := %DB100.DBB47;
END_REGION

REGION Network 14: op_3
   RUNG wire#powerrail
      Move(in := %DB100.DBB64, out1 => %DB100.DBB270)
      Move(in := %DB100.DBB65, out1 => %DB100.DBB271)
   END_RUNG
   RUNG wire#powerrail
      Move(in := %DB100.DBB66, out1 => %DB100.DBB272)
      Move(in := %DB100.DBB67, out1 => %DB100.DBB273)
   END_RUNG
   // the same network as SCL:
   %DB100.DBB270 := %DB100.DBB64;
   %DB100.DBB271 := %DB100.DBB65;
   %DB100.DBB272 := %DB100.DBB66;
   %DB100.DBB273 := %DB100.DBB67;
END_REGION

REGION Network 15 (SCL)
   IF "CONTROL_LINE_DB".trig.reset_error_all = TRUE THEN
       // alarm global
       %DB100. := 0;
       %DB100. := 0;
       // wrong global
       %DB100. := 0;
       %DB100. := 0;
       // op_0
       // alarm
       %DB100. := 0;
       %DB100. := 0;
       // wrong
       %DB100. := 0;
       %DB100. := 0;
       // op_1
       // alarm
       %DB100. := 0;
       %DB100. := 0;
       // wrong
       %DB100. := 0;
       %DB100. := 0;
       // op_2
       // alarm
       %DB100. := 0;
       %DB100. := 0;
       // wrong
       %DB100. := 0;
       %DB100. := 0;
       // op_3
       // alarm
       %DB100. := 0;
       %DB100. := 0;
       // wrong
       %DB100. := 0;
       %DB100. := 0;
       // op_4
       // alarm
       %DB100. := 0;
       %DB100. := 0;
       // wrong
       %DB100. := 0;
       %DB100. := 0;
       // op_5
       // alarm
       %DB100. := 0;
       %DB100. := 0;
       // wrong
       %DB100. := 0;
       %DB100. := 0;
   END_IF;
END_REGION

REGION Network 16 (SCL)
   //"DB_ALARM".op_0_m_0 := "DB_ALARM".OP0.M_0;
   //"DB_ALARM".op_1_m_0 := "DB_ALARM".OP1.M_0;
   //"DB_ALARM".op_2_m_0 := "DB_ALARM".OP2.A1;
   //"DB_ALARM".op_2_m_1 := "DB_ALARM".OP2.A2;
   //"DB_ALARM".op_2_m_2 := "DB_ALARM".OP2.A3;
   //"DB_ALARM".op_2_m_3 := "DB_ALARM".OP2.A4;
   //"DB_ALARM".op_3_m_0 := "DB_ALARM".OP3.B1;
END_REGION
END_FUNCTION

FUNCTION_BLOCK "CONTROL_LINE"   // FB7, LAD
{ S7_Optimized_Access := 'TRUE' }
// stored: MemoryReserve 100, SetENOAutomatically false
   VAR
      TIMER_reset { S7_SetPoint := 'True'} : TON_TIME;
      P_TRIG_INICIAL : Bool;
      P_TRIG_RESET : Bool;
      AUTOMAT { S7_SetPoint := 'True'} : "SENSOR";
      MANUAL { S7_SetPoint := 'True'} : "SENSOR";
      SENSOR_3 { S7_SetPoint := 'True'} : "SENSOR";
      SENSOR_4 { S7_SetPoint := 'True'} : "SENSOR";
      SENSOR_5 { S7_SetPoint := 'True'} : "SENSOR";
      SENSOR_6 { S7_SetPoint := 'True'} : "SENSOR";
      SENSOR_7 { S7_SetPoint := 'True'} : "SENSOR";
      SENSOR_8 { S7_SetPoint := 'True'} : "SENSOR";
      SENSOR_9 { S7_SetPoint := 'True'} : "SENSOR";
      SENSOR_10 { S7_SetPoint := 'True'} : "SENSOR";
      SENSOR_11 { S7_SetPoint := 'True'} : "SENSOR";
      dvere_L_A { S7_SetPoint := 'True'} : "SENSOR";
      dvere_L_B { S7_SetPoint := 'True'} : "SENSOR";
      dvere_P_A { S7_SetPoint := 'True'} : "SENSOR";
      dvere_P_B { S7_SetPoint := 'True'} : "SENSOR";
      SEN_STRUCT : Struct
         AUTOMAT : Bool;
         AUTOMAT_NEG : Bool;
         MANUAL : Bool;
         MANUAL_NEG : Bool;
         SENSOR_TLAKU : Bool;
         SENSOR_TLAKU_NEG : Bool;
         power : Bool;
         power_neg : Bool;
         safety : Bool;
         safety_neg : Bool;
         s_10 : Bool;
         TLA_STOP : Bool;
         TLA_STOP_NEG : Bool;
         TLA_START : Bool;
         TLA_START_NEG : Bool;
         TLA_KVIT : Bool;
         TLA_KVIT_NEG : Bool;
         s_17 : Bool;
         S19 : Bool;
         L1_OK : Bool;
         L1_NOT_OK : Bool;
         L2_OK : Bool;
         L2_NOT_OK : Bool;
         L3_OK : Bool;
         L3_NOT_OK : Bool;
         dvere_L_A : Bool;
         dvere_L_B : Bool;
         dvere_P_A : Bool;
         dvere_P_B : Bool;
         S30 : Bool;
         S31 : Bool;
         LASER_MEMOR : Bool;
      END_STRUCT;
      "M" : Struct
         P_TRIK_hmi_manual : Bool;
         p_trig_hmi_automat : Bool;
         N_TRIG_REZIM : Bool;
         M_4 : Bool;
         hlaseni_chyby : Bool;
         M_6 : Bool;
         M_7 : Bool;
         M_8 : Bool;
         M_9 : Bool;
         p_Trig_al : Bool;
         n_trig_al : Bool;
         p_trig_wro : Bool;
         n_trig_wro : Bool;
         M_14 : Bool;
         M_15 : Bool;
         N_TRIG_MANUAL : Bool;
         M_17 : Bool;
         M_18 : Bool;
         M_19 : Bool;
         M_20 : Bool;
         M_21 : Bool;
         M_22 : Bool;
         M_23 : Bool;
         M_24 : Bool;
         M_25 : Bool;
         M_26 : Bool;
         M_27 : Bool;
         M_28 : Bool;
         M_29 : Bool;
         M_30 : Bool;
         M_31 : Bool;
         M_32 : Bool;
      END_STRUCT;
      trig : Struct
         reset_error_all : Bool;
         TRIG_FOR_OP_4_AUTOMAT : Bool;
         t_3 : Bool;
         t_4 : Bool;
         t_5 : Bool;
         t_6 : Bool;
         t_7 : Bool;
         t_8 : Bool;
      END_STRUCT;
      SQCR : Int;
      job_mailbox : Array[0..3] of Word;
      n_trig_res_auit : Bool;
      inicial_control { S7_SetPoint := 'True'} : TON_TIME;
      SQCR_SAFETY { S7_SetPoint := 'True'} : Int;
      n_trig_RESET_AUT : Bool;
      P_TRIG_RESET_SAFETY : Bool;
      air { S7_SetPoint := 'True'} : TON_TIME;
      HMI_ALARM { S7_SetPoint := 'True'} : Int;
   END_VAR
   VAR_TEMP
      "string" : String;
      smaz_me : Bool;
      majak_green_s1 : Bool;
      majak_red_s1 : Bool;
      majak_yelou_s1 : Bool;
      majak_blue_s1 : Bool;
      majak_orange_s1 : Bool;
      majak_green_s2 : Bool;
      majak_red_s2 : Bool;
      majak_yelou_s2 : Bool;
      majak_blue_s2 : Bool;
      majak_orange_s2 : Bool;
      majak_green_s3 : Bool;
      majak_red_s3 : Bool;
      majak_yelou_s3 : Bool;
      majak_blue_s3 : Bool;
      majak_orange_s3 : Bool;
      majak_green_s4 : Bool;
      majak_red_s4 : Bool;
      majak_yelou_s4 : Bool;
      majak_blue_s4 : Bool;
      majak_orange_s4 : Bool;
      majak_green_s5 : Bool;
      majak_red_s5 : Bool;
      majak_yelou_s5 : Bool;
      majak_blue_s5 : Bool;
      majak_orange_s5 : Bool;
   END_VAR
   VAR CONSTANT
      STEP_0_FIRST_START : Int := 0;
      STEP_3 : Int := 3;
      STEP_5 : Int := 5;
      STEP_10 : Int := 10;
      STEP_15 : Int := 15;
      STEP_20 : Int := 20;
      STEP_25 : Int := 25;
      STEP_27 : Int := 27;
      STEP_30 : Int := 30;
      STEP_35 : Int := 35;
      STEP_40 : Int := 40;
      STEP_45 : Int := 45;
      STEP_48 : Int := 48;
      STEP_50 : Int := 50;
      STEP_52 : Int := 52;
      STEP_55 : Int := 55;
      STEP_60 : Int := 60;
      STEP_65 : Int := 65;
      STEP_70 : Int := 70;
      STEP_75 : Int := 75;
      STEP_80 : Int := 80;
      STEP_85 : Int := 85;
      STEP_90 : Int := 90;
      STEP_95 : Int := 95;
      STEP_100 : Int := 100;
      STEO_105 : Int := 105;
   END_VAR
   VAR_TEMP   // added for the SCL form of the ladder/FBD networks
      _w1 : Bool;
      _w2 : Bool;
      _w3 : Bool;
      _w4 : Bool;
      _w5 : Bool;
   END_VAR
BEGIN

REGION Network 1 (SCL)
   // SET  BASIC ELEMENTS
   // odpojení nepoužívaných kontaktů
   "LOG_0" := 0;
   "LOG_1" := 1;
   "SMAZ_ME_0" := 0;
   "SMAZ_ME_1" := 1;
END_REGION

REGION Network 2: SENSORS
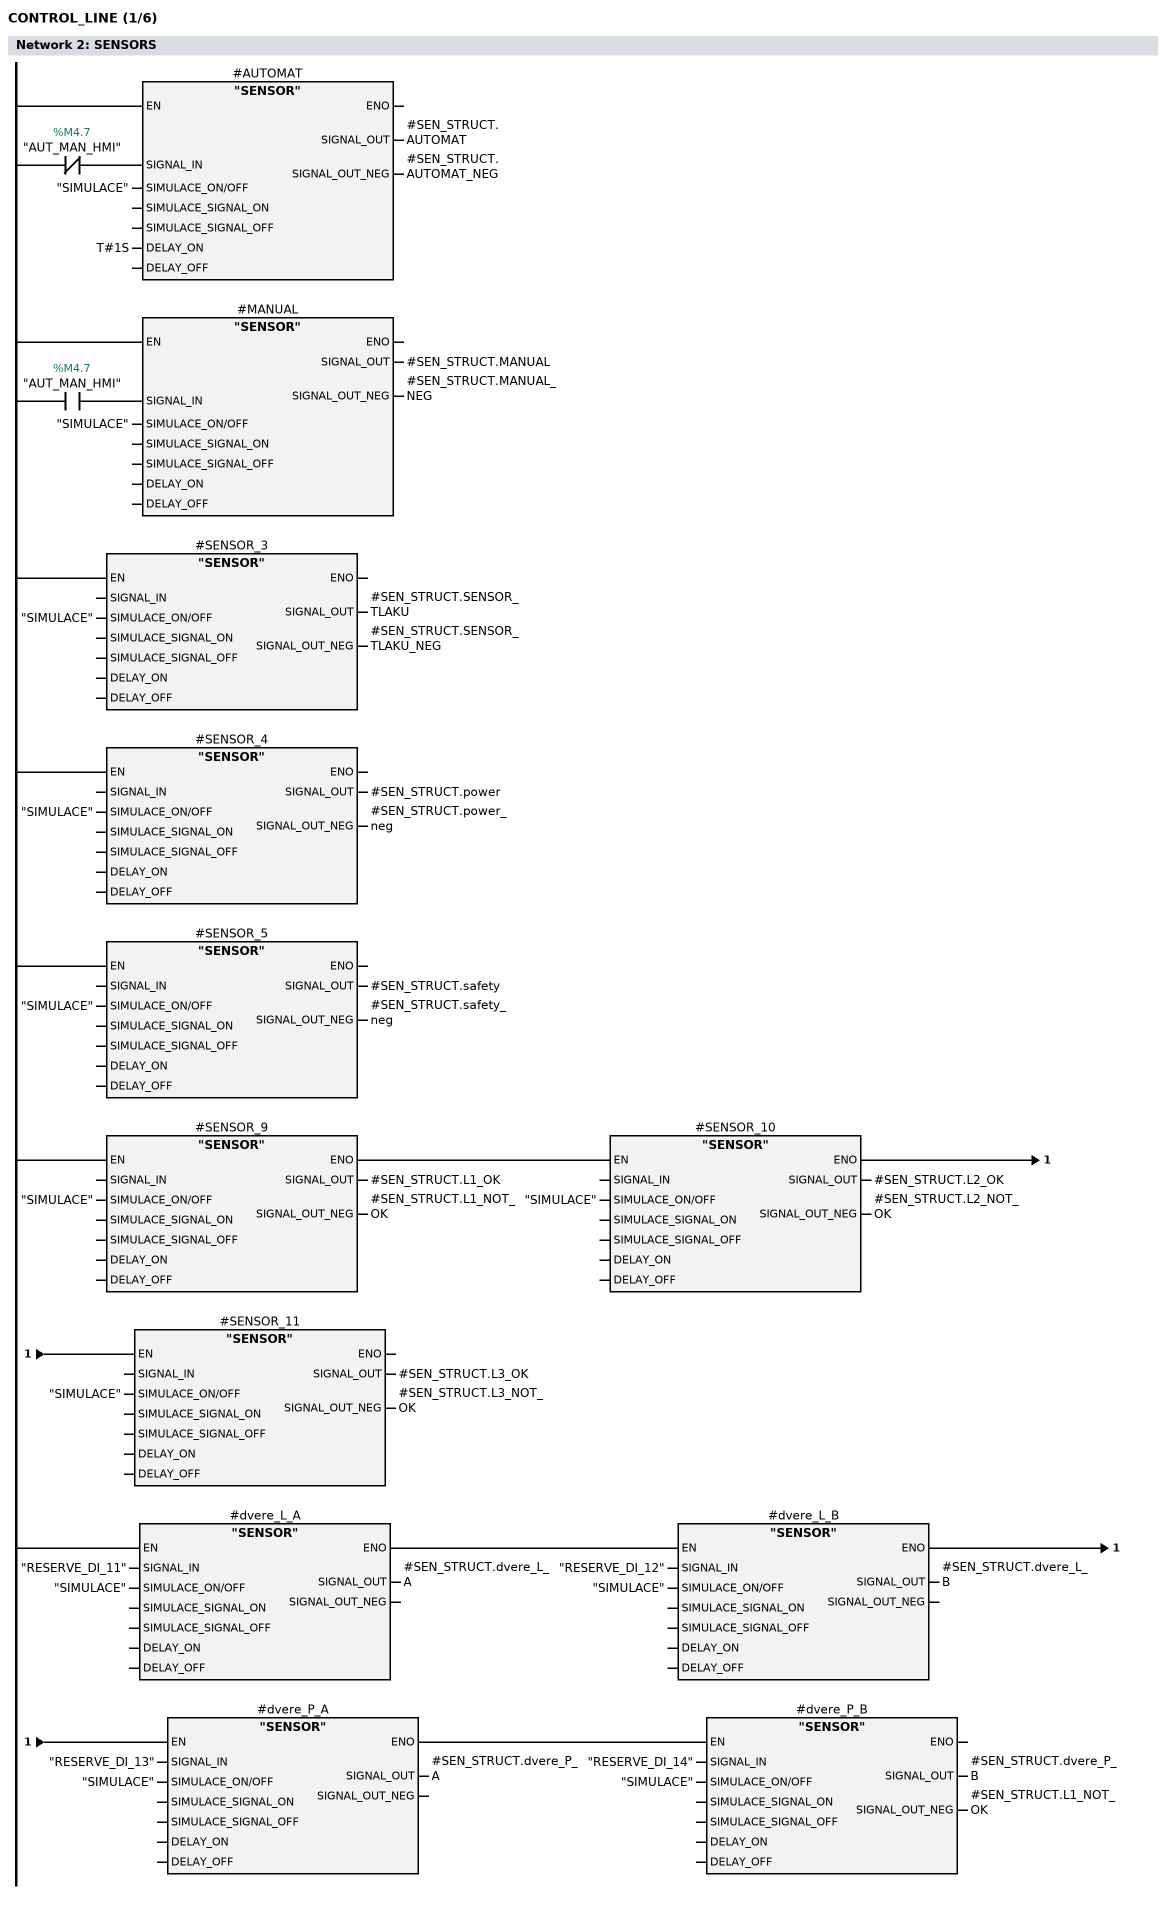
   RUNG wire#powerrail
      #AUTOMAT(SIGNAL_IN := wire#w1, "SIMULACE_ON/OFF" := "SIMULACE", SIMULACE_SIGNAL_ON :=, SIMULACE_SIGNAL_OFF :=, DELAY_ON := T#1S, DELAY_OFF :=, SIGNAL_OUT => #SEN_STRUCT.AUTOMAT, SIGNAL_OUT_NEG => #SEN_STRUCT.AUTOMAT_NEG)
   END_RUNG
   RUNG wire#powerrail
      I_Contact( "AUT_MAN_HMI" )
   END_RUNG wire#w1
   RUNG wire#powerrail
      #MANUAL(SIGNAL_IN := wire#w2, "SIMULACE_ON/OFF" := "SIMULACE", SIMULACE_SIGNAL_ON :=, SIMULACE_SIGNAL_OFF :=, DELAY_ON :=, DELAY_OFF :=, SIGNAL_OUT => #SEN_STRUCT.MANUAL, SIGNAL_OUT_NEG => #SEN_STRUCT.MANUAL_NEG)
   END_RUNG
   RUNG wire#powerrail
      Contact( "AUT_MAN_HMI" )
   END_RUNG wire#w2
   RUNG wire#powerrail
      #SENSOR_3(SIGNAL_IN :=, "SIMULACE_ON/OFF" := "SIMULACE", SIMULACE_SIGNAL_ON :=, SIMULACE_SIGNAL_OFF :=, DELAY_ON :=, DELAY_OFF :=, SIGNAL_OUT => #SEN_STRUCT.SENSOR_TLAKU, SIGNAL_OUT_NEG => #SEN_STRUCT.SENSOR_TLAKU_NEG)
   END_RUNG
   RUNG wire#powerrail
      #SENSOR_4(SIGNAL_IN :=, "SIMULACE_ON/OFF" := "SIMULACE", SIMULACE_SIGNAL_ON :=, SIMULACE_SIGNAL_OFF :=, DELAY_ON :=, DELAY_OFF :=, SIGNAL_OUT => #SEN_STRUCT.power, SIGNAL_OUT_NEG => #SEN_STRUCT.power_neg)
   END_RUNG
   RUNG wire#powerrail
      #SENSOR_5(SIGNAL_IN :=, "SIMULACE_ON/OFF" := "SIMULACE", SIMULACE_SIGNAL_ON :=, SIMULACE_SIGNAL_OFF :=, DELAY_ON :=, DELAY_OFF :=, SIGNAL_OUT => #SEN_STRUCT.safety, SIGNAL_OUT_NEG => #SEN_STRUCT.safety_neg)
   END_RUNG
   RUNG wire#powerrail
      #SENSOR_9(SIGNAL_IN :=, "SIMULACE_ON/OFF" := "SIMULACE", SIMULACE_SIGNAL_ON :=, SIMULACE_SIGNAL_OFF :=, DELAY_ON :=, DELAY_OFF :=, SIGNAL_OUT => #SEN_STRUCT.L1_OK, SIGNAL_OUT_NEG => #SEN_STRUCT.L1_NOT_OK)
      #SENSOR_10(SIGNAL_IN :=, "SIMULACE_ON/OFF" := "SIMULACE", SIMULACE_SIGNAL_ON :=, SIMULACE_SIGNAL_OFF :=, DELAY_ON :=, DELAY_OFF :=, SIGNAL_OUT => #SEN_STRUCT.L2_OK, SIGNAL_OUT_NEG => #SEN_STRUCT.L2_NOT_OK)
      #SENSOR_11(SIGNAL_IN :=, "SIMULACE_ON/OFF" := "SIMULACE", SIMULACE_SIGNAL_ON :=, SIMULACE_SIGNAL_OFF :=, DELAY_ON :=, DELAY_OFF :=, SIGNAL_OUT => #SEN_STRUCT.L3_OK, SIGNAL_OUT_NEG => #SEN_STRUCT.L3_NOT_OK)
   END_RUNG
   RUNG wire#powerrail
      #dvere_L_A(SIGNAL_IN := "RESERVE_DI_11", "SIMULACE_ON/OFF" := "SIMULACE", SIMULACE_SIGNAL_ON :=, SIMULACE_SIGNAL_OFF :=, DELAY_ON :=, DELAY_OFF :=, SIGNAL_OUT => #SEN_STRUCT.dvere_L_A, SIGNAL_OUT_NEG =>)
      #dvere_L_B(SIGNAL_IN := "RESERVE_DI_12", "SIMULACE_ON/OFF" := "SIMULACE", SIMULACE_SIGNAL_ON :=, SIMULACE_SIGNAL_OFF :=, DELAY_ON :=, DELAY_OFF :=, SIGNAL_OUT => #SEN_STRUCT.dvere_L_B, SIGNAL_OUT_NEG =>)
      #dvere_P_A(SIGNAL_IN := "RESERVE_DI_13", "SIMULACE_ON/OFF" := "SIMULACE", SIMULACE_SIGNAL_ON :=, SIMULACE_SIGNAL_OFF :=, DELAY_ON :=, DELAY_OFF :=, SIGNAL_OUT => #SEN_STRUCT.dvere_P_A, SIGNAL_OUT_NEG =>)
      #dvere_P_B(SIGNAL_IN := "RESERVE_DI_14", "SIMULACE_ON/OFF" := "SIMULACE", SIMULACE_SIGNAL_ON :=, SIMULACE_SIGNAL_OFF :=, DELAY_ON :=, DELAY_OFF :=, SIGNAL_OUT => #SEN_STRUCT.dvere_P_B, SIGNAL_OUT_NEG => #SEN_STRUCT.L1_NOT_OK)
   END_RUNG
   // the same network as SCL:
   #AUTOMAT(SIGNAL_IN := NOT "AUT_MAN_HMI",   // "SENSOR"
            "SIMULACE_ON/OFF" := "SIMULACE",
            DELAY_ON := T#1S,
            SIGNAL_OUT => #SEN_STRUCT.AUTOMAT,
            SIGNAL_OUT_NEG => #SEN_STRUCT.AUTOMAT_NEG);
   #MANUAL(SIGNAL_IN := "AUT_MAN_HMI",   // "SENSOR"
           "SIMULACE_ON/OFF" := "SIMULACE",
           SIGNAL_OUT => #SEN_STRUCT.MANUAL,
           SIGNAL_OUT_NEG => #SEN_STRUCT.MANUAL_NEG);
   #SENSOR_3("SIMULACE_ON/OFF" := "SIMULACE",   // "SENSOR"
             SIGNAL_OUT => #SEN_STRUCT.SENSOR_TLAKU,
             SIGNAL_OUT_NEG => #SEN_STRUCT.SENSOR_TLAKU_NEG);
   #SENSOR_4("SIMULACE_ON/OFF" := "SIMULACE",   // "SENSOR"
             SIGNAL_OUT => #SEN_STRUCT.power,
             SIGNAL_OUT_NEG => #SEN_STRUCT.power_neg);
   #SENSOR_5("SIMULACE_ON/OFF" := "SIMULACE",   // "SENSOR"
             SIGNAL_OUT => #SEN_STRUCT.safety,
             SIGNAL_OUT_NEG => #SEN_STRUCT.safety_neg);
   #SENSOR_9("SIMULACE_ON/OFF" := "SIMULACE",   // "SENSOR"
             SIGNAL_OUT => #SEN_STRUCT.L1_OK,
             SIGNAL_OUT_NEG => #SEN_STRUCT.L1_NOT_OK,
             ENO => #_w1);
   #SENSOR_10(EN := #_w1,   // "SENSOR"
              "SIMULACE_ON/OFF" := "SIMULACE",
              SIGNAL_OUT => #SEN_STRUCT.L2_OK,
              SIGNAL_OUT_NEG => #SEN_STRUCT.L2_NOT_OK,
              ENO => #_w2);
   IF #_w2 THEN
       #SENSOR_11("SIMULACE_ON/OFF" := "SIMULACE",   // "SENSOR"
                  SIGNAL_OUT => #SEN_STRUCT.L3_OK,
                  SIGNAL_OUT_NEG => #SEN_STRUCT.L3_NOT_OK);
   END_IF;
   #dvere_L_A(SIGNAL_IN := "RESERVE_DI_11",   // "SENSOR"
              "SIMULACE_ON/OFF" := "SIMULACE",
              SIGNAL_OUT => #SEN_STRUCT.dvere_L_A,
              ENO => #_w3);
   #dvere_L_B(EN := #_w3,   // "SENSOR"
              SIGNAL_IN := "RESERVE_DI_12",
              "SIMULACE_ON/OFF" := "SIMULACE",
              SIGNAL_OUT => #SEN_STRUCT.dvere_L_B,
              ENO => #_w4);
   #dvere_P_A(EN := #_w4,   // "SENSOR"
              SIGNAL_IN := "RESERVE_DI_13",
              "SIMULACE_ON/OFF" := "SIMULACE",
              SIGNAL_OUT => #SEN_STRUCT.dvere_P_A,
              ENO => #_w5);
   IF #_w5 THEN
       #dvere_P_B(SIGNAL_IN := "RESERVE_DI_14",   // "SENSOR"
                  "SIMULACE_ON/OFF" := "SIMULACE",
                  SIGNAL_OUT => #SEN_STRUCT.dvere_P_B,
                  SIGNAL_OUT_NEG => #SEN_STRUCT.L1_NOT_OK);
   END_IF;
END_REGION

REGION Network 3 (SCL): ALARMY OP1/OP2 -> HMI
   // ===== ALARMY -> HMI (DB_ALARM.alarm_line, HMI ID 1-16) =====
   // bit 9 (ID 10 aplikator) a bit 14 (ID 15 tlak vzduchu) = firemni standard, nepouzivat

   // bit 0 - tiskarna nekomunikuje (OP2 se nevrati do kroku 5 do 15 s)
   "DB_ALARM".T_tiskarna.TON(IN := "AUTOMAT" AND "OP2_DB".SQCR <> 5,
                             PT := T#15S);
   "DB_ALARM".alarm_line.%X0 := "DB_ALARM".T_tiskarna.Q;

   // bity 1-3 - kamery offline (jen v automatu)
   "DB_ALARM".alarm_line.%X1 := "AUTOMAT" AND NOT "COG_FOLIE_L_is3800-Online";
   "DB_ALARM".alarm_line.%X2 := "AUTOMAT" AND NOT "COG_FOLIE_P_is3800-Online";
   "DB_ALARM".alarm_line.%X3 := "AUTOMAT" AND NOT "COG_ETIKETA_is3800-Online"
   AND NOT "OP1_DB".Kam_Etiketa_Job.aktivni;   // pri loadu jobu je kamera chvili offline

   // bit 4 - chybne datum v recepture
   "DB_ALARM".alarm_line.%X4 := "OP2_DB".Tisk.datum_chyba;

   // bit 5 - fronta plna
   "DB_ALARM".alarm_line.%X5 := "OP1_DB".Kamera.fronta_plna;

   // bit 6 - job horni kamery se nenacetl
   //"DB_ALARM".alarm_line.%X6 := "OP1_DB".Kam_Etiketa_Job.chyba;

   // bity 7-8 - otevrene dvere (signaly ze site "alarmy")
   "DB_ALARM".alarm_line.%X7 := "DB_ALARM".WRONG.dvere_L_tevreny;
   "DB_ALARM".alarm_line.%X8 := "DB_ALARM".WRONG.dvere_P_otevreny;

   // souhrnny alarm -> KA19 blika, HMI_ALARM = 10
   "alrm_global" := "DB_ALARM".alarm_line <> 0;
   "DB_ALARM".ALARM.ALARM_GLOBAL := "alrm_global";
END_REGION

REGION Network 4: alarmy
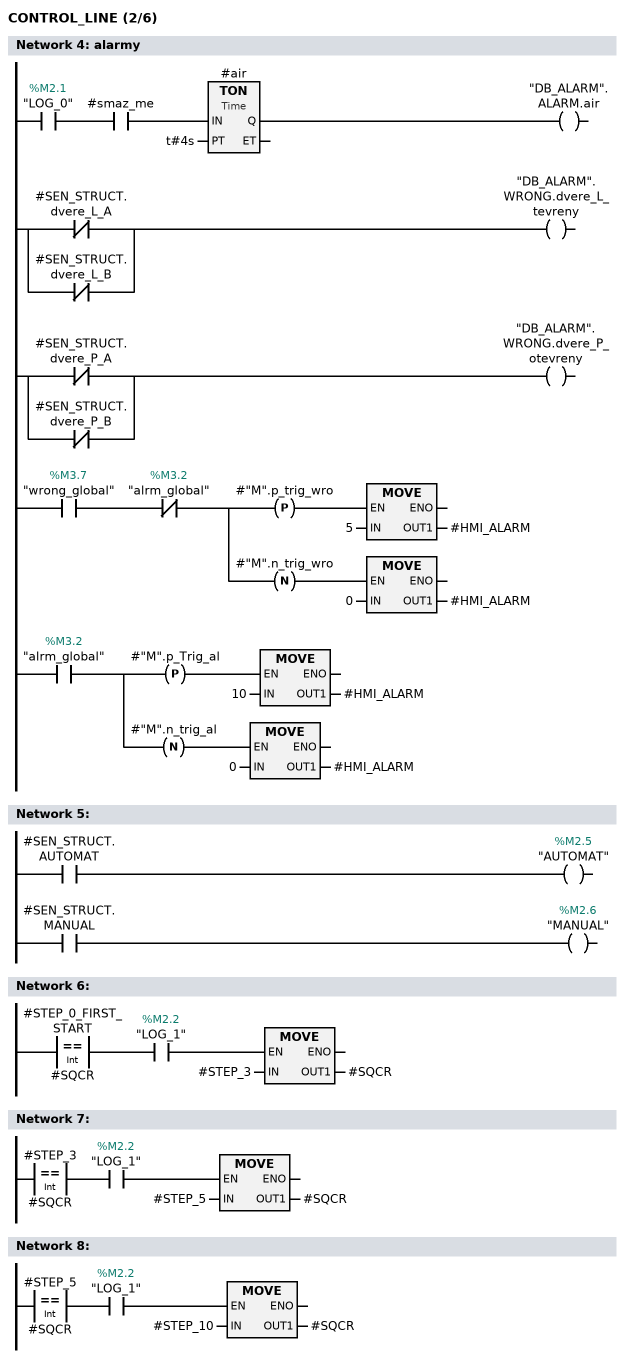
   RUNG wire#powerrail
      Contact( "LOG_0" )
      Contact( #smaz_me )
      { S7_Templates := "time_type := Time" } #air.TON(pt := t#4s, et =>)
      Coil( "DB_ALARM".ALARM.air )
   END_RUNG
   RUNG wire#powerrail
      I_Contact( #SEN_STRUCT.dvere_L_A )
      wire#w1
      Coil( "DB_ALARM".WRONG.dvere_L_tevreny )
   END_RUNG
   RUNG wire#powerrail
      I_Contact( #SEN_STRUCT.dvere_L_B )
   END_RUNG wire#w1
   RUNG wire#powerrail
      I_Contact( #SEN_STRUCT.dvere_P_A )
      wire#w2
      Coil( "DB_ALARM".WRONG.dvere_P_otevreny )
   END_RUNG
   RUNG wire#powerrail
      I_Contact( #SEN_STRUCT.dvere_P_B )
   END_RUNG wire#w2
   RUNG wire#powerrail
      Contact( "wrong_global" )
      I_Contact( "alrm_global" )
      wire#w3
      P_Trig( #"M".p_trig_wro )
      Move(in := 5, out1 => #HMI_ALARM)
   END_RUNG
   RUNG wire#w3
      N_Trig( #"M".n_trig_wro )
      Move(in := 0, out1 => #HMI_ALARM)
   END_RUNG
   RUNG wire#powerrail
      Contact( "alrm_global" )
      wire#w4
      P_Trig( #"M".p_Trig_al )
      Move(in := 10, out1 => #HMI_ALARM)
   END_RUNG
   RUNG wire#w4
      N_Trig( #"M".n_trig_al )
      Move(in := 0, out1 => #HMI_ALARM)
   END_RUNG
   // the same network as SCL:
   #air(IN := "LOG_0" AND #smaz_me, PT := t#4s);   // TON
   "DB_ALARM".ALARM.air := #air.Q;
   "DB_ALARM".WRONG.dvere_L_tevreny := NOT #SEN_STRUCT.dvere_L_A OR NOT #SEN_STRUCT.dvere_L_B;
   "DB_ALARM".WRONG.dvere_P_otevreny := NOT #SEN_STRUCT.dvere_P_A OR NOT #SEN_STRUCT.dvere_P_B;
   #_w1 := "wrong_global" AND NOT "alrm_global";
   #_w2 := #_w1 AND NOT #"M".p_trig_wro;   // rising edge
   #"M".p_trig_wro := #_w1;
   IF #_w2 THEN #HMI_ALARM := 5; END_IF;
   #_w3 := NOT #_w1 AND #"M".n_trig_wro;   // falling edge
   #"M".n_trig_wro := #_w1;
   IF #_w3 THEN #HMI_ALARM := 0; END_IF;
   #_w4 := "alrm_global" AND NOT #"M".p_Trig_al;   // rising edge
   #"M".p_Trig_al := "alrm_global";
   IF #_w4 THEN #HMI_ALARM := 10; END_IF;
   #_w5 := NOT "alrm_global" AND #"M".n_trig_al;   // falling edge
   #"M".n_trig_al := "alrm_global";
   IF #_w5 THEN #HMI_ALARM := 0; END_IF;
END_REGION

REGION Network 5
   RUNG wire#powerrail
      Contact( #SEN_STRUCT.AUTOMAT )
      Coil( "AUTOMAT" )
   END_RUNG
   RUNG wire#powerrail
      Contact( #SEN_STRUCT.MANUAL )
      Coil( "MANUAL" )
   END_RUNG
   // the same network as SCL:
   "AUTOMAT" := #SEN_STRUCT.AUTOMAT;
   "MANUAL" := #SEN_STRUCT.MANUAL;
END_REGION

REGION Network 6
   RUNG wire#powerrail
      { S7_Templates := "SrcType := Int" } EQ_Contact(in1 := #STEP_0_FIRST_START, in2 := #SQCR)
      Contact( "LOG_1" )
      Move(in := #STEP_3, out1 => #SQCR)
   END_RUNG
   // the same network as SCL:
   IF (#STEP_0_FIRST_START = #SQCR) AND "LOG_1" THEN #SQCR := #STEP_3; END_IF;
END_REGION

REGION Network 7
   RUNG wire#powerrail
      { S7_Templates := "SrcType := Int" } EQ_Contact(in1 := #STEP_3, in2 := #SQCR)
      Contact( "LOG_1" )
      Move(in := #STEP_5, out1 => #SQCR)
   END_RUNG
   // the same network as SCL:
   IF (#STEP_3 = #SQCR) AND "LOG_1" THEN #SQCR := #STEP_5; END_IF;
END_REGION

REGION Network 8
   RUNG wire#powerrail
      { S7_Templates := "SrcType := Int" } EQ_Contact(in1 := #STEP_5, in2 := #SQCR)
      Contact( "LOG_1" )
      Move(in := #STEP_10, out1 => #SQCR)
   END_RUNG
   // the same network as SCL:
   IF (#STEP_5 = #SQCR) AND "LOG_1" THEN #SQCR := #STEP_10; END_IF;
END_REGION

REGION Network 9
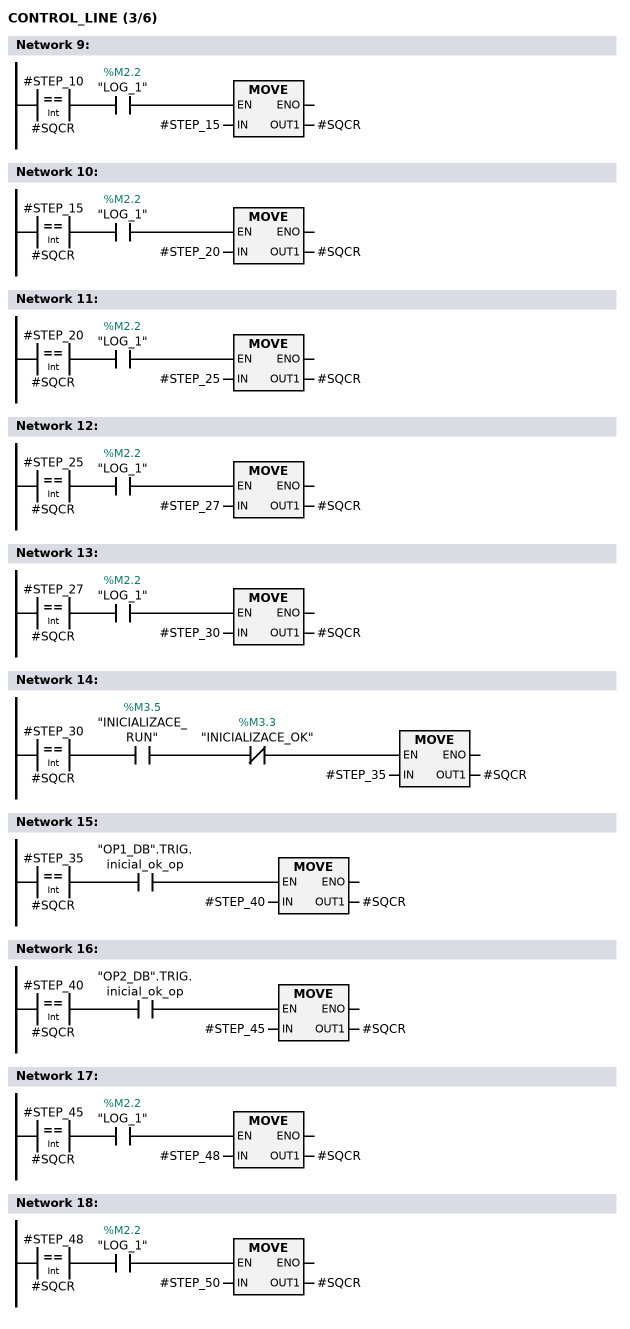
   RUNG wire#powerrail
      { S7_Templates := "SrcType := Int" } EQ_Contact(in1 := #STEP_10, in2 := #SQCR)
      Contact( "LOG_1" )
      Move(in := #STEP_15, out1 => #SQCR)
   END_RUNG
   // the same network as SCL:
   IF (#STEP_10 = #SQCR) AND "LOG_1" THEN #SQCR := #STEP_15; END_IF;
END_REGION

REGION Network 10
   RUNG wire#powerrail
      { S7_Templates := "SrcType := Int" } EQ_Contact(in1 := #STEP_15, in2 := #SQCR)
      Contact( "LOG_1" )
      Move(in := #STEP_20, out1 => #SQCR)
   END_RUNG
   // the same network as SCL:
   IF (#STEP_15 = #SQCR) AND "LOG_1" THEN #SQCR := #STEP_20; END_IF;
END_REGION

REGION Network 11
   RUNG wire#powerrail
      { S7_Templates := "SrcType := Int" } EQ_Contact(in1 := #STEP_20, in2 := #SQCR)
      Contact( "LOG_1" )
      Move(in := #STEP_25, out1 => #SQCR)
   END_RUNG
   // the same network as SCL:
   IF (#STEP_20 = #SQCR) AND "LOG_1" THEN #SQCR := #STEP_25; END_IF;
END_REGION

REGION Network 12
   RUNG wire#powerrail
      { S7_Templates := "SrcType := Int" } EQ_Contact(in1 := #STEP_25, in2 := #SQCR)
      Contact( "LOG_1" )
      Move(in := #STEP_27, out1 => #SQCR)
   END_RUNG
   // the same network as SCL:
   IF (#STEP_25 = #SQCR) AND "LOG_1" THEN #SQCR := #STEP_27; END_IF;
END_REGION

REGION Network 13
   RUNG wire#powerrail
      { S7_Templates := "SrcType := Int" } EQ_Contact(in1 := #STEP_27, in2 := #SQCR)
      Contact( "LOG_1" )
      Move(in := #STEP_30, out1 => #SQCR)
   END_RUNG
   // the same network as SCL:
   IF (#STEP_27 = #SQCR) AND "LOG_1" THEN #SQCR := #STEP_30; END_IF;
END_REGION

REGION Network 14
   RUNG wire#powerrail
      { S7_Templates := "SrcType := Int" } EQ_Contact(in1 := #STEP_30, in2 := #SQCR)
      Contact( "INICIALIZACE_RUN" )
      I_Contact( "INICIALIZACE_OK" )
      Move(in := #STEP_35, out1 => #SQCR)
   END_RUNG
   // the same network as SCL:
   IF (#STEP_30 = #SQCR) AND "INICIALIZACE_RUN" AND NOT "INICIALIZACE_OK" THEN #SQCR := #STEP_35; END_IF;
END_REGION

REGION Network 15
   RUNG wire#powerrail
      { S7_Templates := "SrcType := Int" } EQ_Contact(in1 := #STEP_35, in2 := #SQCR)
      Contact( "OP1_DB".TRIG.inicial_ok_op )
      Move(in := #STEP_40, out1 => #SQCR)
   END_RUNG
   // the same network as SCL:
   IF (#STEP_35 = #SQCR) AND "OP1_DB".TRIG.inicial_ok_op THEN #SQCR := #STEP_40; END_IF;
END_REGION

REGION Network 16
   RUNG wire#powerrail
      { S7_Templates := "SrcType := Int" } EQ_Contact(in1 := #STEP_40, in2 := #SQCR)
      Contact( "OP2_DB".TRIG.inicial_ok_op )
      Move(in := #STEP_45, out1 => #SQCR)
   END_RUNG
   // the same network as SCL:
   IF (#STEP_40 = #SQCR) AND "OP2_DB".TRIG.inicial_ok_op THEN #SQCR := #STEP_45; END_IF;
END_REGION

REGION Network 17
   RUNG wire#powerrail
      { S7_Templates := "SrcType := Int" } EQ_Contact(in1 := #STEP_45, in2 := #SQCR)
      Contact( "LOG_1" )
      Move(in := #STEP_48, out1 => #SQCR)
   END_RUNG
   // the same network as SCL:
   IF (#STEP_45 = #SQCR) AND "LOG_1" THEN #SQCR := #STEP_48; END_IF;
END_REGION

REGION Network 18
   RUNG wire#powerrail
      { S7_Templates := "SrcType := Int" } EQ_Contact(in1 := #STEP_48, in2 := #SQCR)
      Contact( "LOG_1" )
      Move(in := #STEP_50, out1 => #SQCR)
   END_RUNG
   // the same network as SCL:
   IF (#STEP_48 = #SQCR) AND "LOG_1" THEN #SQCR := #STEP_50; END_IF;
END_REGION

REGION Network 19
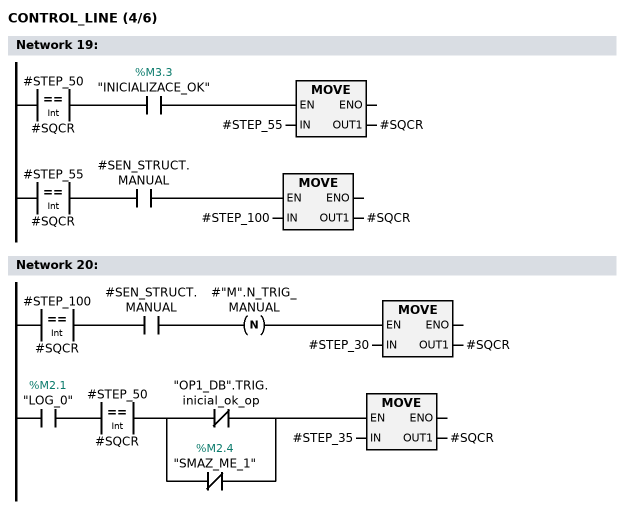
   RUNG wire#powerrail
      { S7_Templates := "SrcType := Int" } EQ_Contact(in1 := #STEP_50, in2 := #SQCR)
      Contact( "INICIALIZACE_OK" )
      Move(in := #STEP_55, out1 => #SQCR)
   END_RUNG
   RUNG wire#powerrail
      { S7_Templates := "SrcType := Int" } EQ_Contact(in1 := #STEP_55, in2 := #SQCR)
      Contact( #SEN_STRUCT.MANUAL )
      Move(in := #STEP_100, out1 => #SQCR)
   END_RUNG
   // the same network as SCL:
   IF (#STEP_50 = #SQCR) AND "INICIALIZACE_OK" THEN #SQCR := #STEP_55; END_IF;
   IF (#STEP_55 = #SQCR) AND #SEN_STRUCT.MANUAL THEN #SQCR := #STEP_100; END_IF;
END_REGION

REGION Network 20
   RUNG wire#powerrail
      { S7_Templates := "SrcType := Int" } EQ_Contact(in1 := #STEP_100, in2 := #SQCR)
      Contact( #SEN_STRUCT.MANUAL )
      N_Trig( #"M".N_TRIG_MANUAL )
      Move(in := #STEP_30, out1 => #SQCR)
   END_RUNG
   RUNG wire#powerrail
      Contact( "LOG_0" )
      { S7_Templates := "SrcType := Int" } EQ_Contact(in1 := #STEP_50, in2 := #SQCR)
      wire#w1
      I_Contact( "OP1_DB".TRIG.inicial_ok_op )
      wire#w2
      Move(in := #STEP_35, out1 => #SQCR)
   END_RUNG
   RUNG wire#w1
      I_Contact( "SMAZ_ME_1" )
   END_RUNG wire#w2
   // the same network as SCL:
   #_w1 := (#STEP_100 = #SQCR) AND #SEN_STRUCT.MANUAL;
   #_w2 := NOT #_w1 AND #"M".N_TRIG_MANUAL;   // falling edge
   #"M".N_TRIG_MANUAL := #_w1;
   IF #_w2 THEN #SQCR := #STEP_30; END_IF;
   IF "LOG_0" AND (#STEP_50 = #SQCR) AND (NOT "OP1_DB".TRIG.inicial_ok_op OR NOT "SMAZ_ME_1") THEN
       #SQCR := #STEP_35;
   END_IF;
END_REGION

REGION Network 21: LEDKY
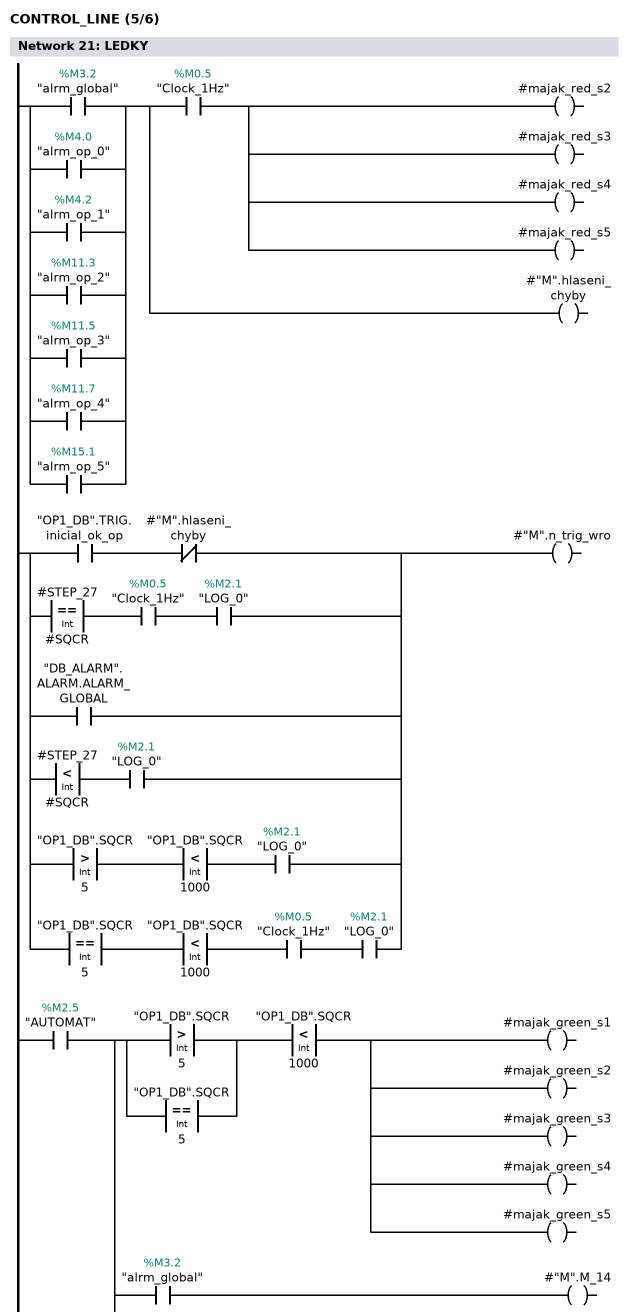
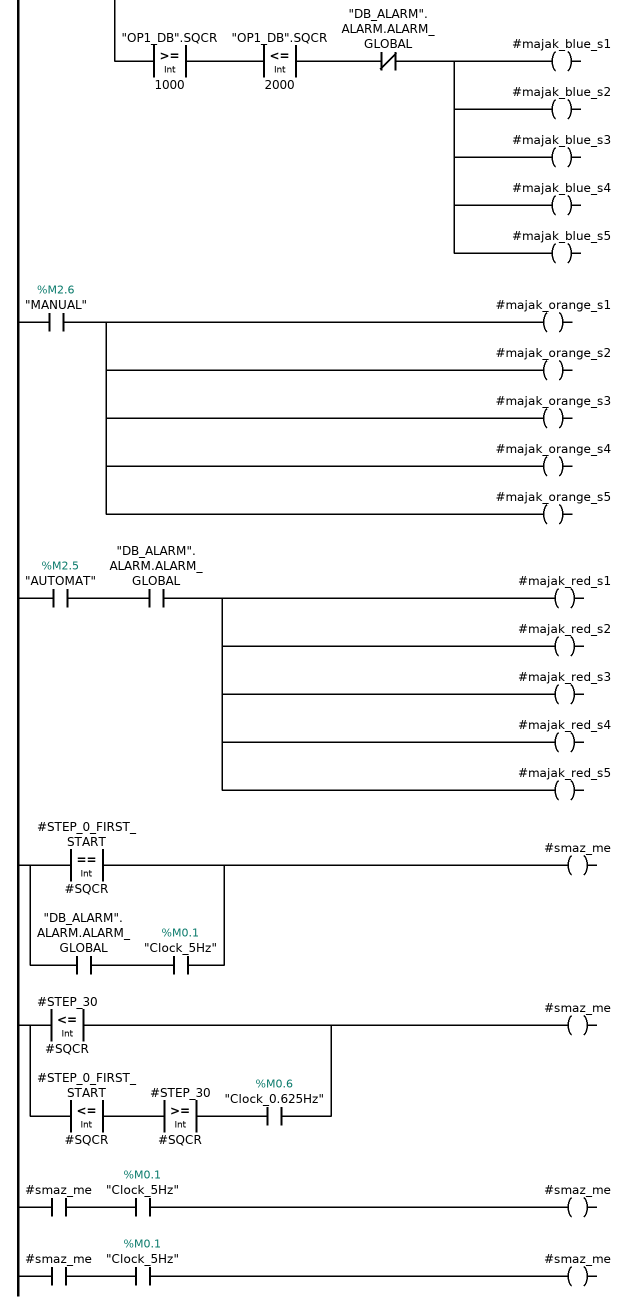
   RUNG wire#powerrail
      Contact( "alrm_global" )
      wire#w1
      Contact( "Clock_1Hz" )
      wire#w2
      Coil( #majak_red_s2 )
   END_RUNG
   RUNG wire#powerrail
      Contact( "alrm_op_0" )
   END_RUNG wire#w1
   RUNG wire#powerrail
      Contact( "alrm_op_1" )
   END_RUNG wire#w1
   RUNG wire#powerrail
      Contact( "alrm_op_2" )
   END_RUNG wire#w1
   RUNG wire#powerrail
      Contact( "alrm_op_3" )
   END_RUNG wire#w1
   RUNG wire#powerrail
      Contact( "alrm_op_4" )
   END_RUNG wire#w1
   RUNG wire#powerrail
      Contact( "alrm_op_5" )
   END_RUNG wire#w1
   RUNG wire#w2
      Coil( #majak_red_s3 )
   END_RUNG
   RUNG wire#w2
      Coil( #majak_red_s4 )
   END_RUNG
   RUNG wire#w2
      Coil( #majak_red_s5 )
   END_RUNG
   RUNG wire#w1
      Coil( #"M".hlaseni_chyby )
   END_RUNG
   RUNG wire#powerrail
      Contact( "OP1_DB".TRIG.inicial_ok_op )
      I_Contact( #"M".hlaseni_chyby )
      wire#w3
      Coil( #"M".n_trig_wro )
   END_RUNG
   RUNG wire#powerrail
      { S7_Templates := "SrcType := Int" } EQ_Contact(in1 := #STEP_27, in2 := #SQCR)
      Contact( "Clock_1Hz" )
      Contact( "LOG_0" )
   END_RUNG wire#w3
   RUNG wire#powerrail
      Contact( "DB_ALARM".ALARM.ALARM_GLOBAL )
   END_RUNG wire#w3
   RUNG wire#powerrail
      { S7_Templates := "SrcType := Int" } LT_Contact(in1 := #STEP_27, in2 := #SQCR)
      Contact( "LOG_0" )
   END_RUNG wire#w3
   RUNG wire#powerrail
      { S7_Templates := "SrcType := Int" } GT_Contact(in1 := "OP1_DB".SQCR, in2 := 5)
      { S7_Templates := "SrcType := Int" } LT_Contact(in1 := "OP1_DB".SQCR, in2 := 1000)
      Contact( "LOG_0" )
   END_RUNG wire#w3
   RUNG wire#powerrail
      { S7_Templates := "SrcType := Int" } EQ_Contact(in1 := "OP1_DB".SQCR, in2 := 5)
      { S7_Templates := "SrcType := Int" } LT_Contact(in1 := "OP1_DB".SQCR, in2 := 1000)
      Contact( "Clock_1Hz" )
      Contact( "LOG_0" )
   END_RUNG wire#w3
   RUNG wire#powerrail
      Contact( "AUTOMAT" )
      wire#w4
      { S7_Templates := "SrcType := Int" } GT_Contact(in1 := "OP1_DB".SQCR, in2 := 5)
      wire#w5
      { S7_Templates := "SrcType := Int" } LT_Contact(in1 := "OP1_DB".SQCR, in2 := 1000)
      wire#w6
      Coil( #majak_green_s1 )
   END_RUNG
   RUNG wire#w4
      { S7_Templates := "SrcType := Int" } EQ_Contact(in1 := "OP1_DB".SQCR, in2 := 5)
   END_RUNG wire#w5
   RUNG wire#w6
      Coil( #majak_green_s2 )
   END_RUNG
   RUNG wire#w6
      Coil( #majak_green_s3 )
   END_RUNG
   RUNG wire#w6
      Coil( #majak_green_s4 )
   END_RUNG
   RUNG wire#w6
      Coil( #majak_green_s5 )
   END_RUNG
   RUNG wire#w4
      Contact( "alrm_global" )
      Coil( #"M".M_14 )
   END_RUNG
   RUNG wire#w4
      { S7_Templates := "SrcType := Int" } GE_Contact(in1 := "OP1_DB".SQCR, in2 := 1000)
      { S7_Templates := "SrcType := Int" } LE_Contact(in1 := "OP1_DB".SQCR, in2 := 2000)
      I_Contact( "DB_ALARM".ALARM.ALARM_GLOBAL )
      wire#w7
      Coil( #majak_blue_s1 )
   END_RUNG
   RUNG wire#w7
      Coil( #majak_blue_s2 )
   END_RUNG
   RUNG wire#w7
      Coil( #majak_blue_s3 )
   END_RUNG
   RUNG wire#w7
      Coil( #majak_blue_s4 )
   END_RUNG
   RUNG wire#w7
      Coil( #majak_blue_s5 )
   END_RUNG
   RUNG wire#powerrail
      Contact( "MANUAL" )
      wire#w8
      Coil( #majak_orange_s1 )
   END_RUNG
   RUNG wire#w8
      Coil( #majak_orange_s2 )
   END_RUNG
   RUNG wire#w8
      Coil( #majak_orange_s3 )
   END_RUNG
   RUNG wire#w8
      Coil( #majak_orange_s4 )
   END_RUNG
   RUNG wire#w8
      Coil( #majak_orange_s5 )
   END_RUNG
   RUNG wire#powerrail
      Contact( "AUTOMAT" )
      Contact( "DB_ALARM".ALARM.ALARM_GLOBAL )
      wire#w9
      Coil( #majak_red_s1 )
   END_RUNG
   RUNG wire#w9
      Coil( #majak_red_s2 )
   END_RUNG
   RUNG wire#w9
      Coil( #majak_red_s3 )
   END_RUNG
   RUNG wire#w9
      Coil( #majak_red_s4 )
   END_RUNG
   RUNG wire#w9
      Coil( #majak_red_s5 )
   END_RUNG
   RUNG wire#powerrail
      { S7_Templates := "SrcType := Int" } EQ_Contact(in1 := #STEP_0_FIRST_START, in2 := #SQCR)
      wire#w10
      Coil( #smaz_me )
   END_RUNG
   RUNG wire#powerrail
      Contact( "DB_ALARM".ALARM.ALARM_GLOBAL )
      Contact( "Clock_5Hz" )
   END_RUNG wire#w10
   RUNG wire#powerrail
      { S7_Templates := "SrcType := Int" } LE_Contact(in1 := #STEP_30, in2 := #SQCR)
      wire#w11
      Coil( #smaz_me )
   END_RUNG
   RUNG wire#powerrail
      { S7_Templates := "SrcType := Int" } LE_Contact(in1 := #STEP_0_FIRST_START, in2 := #SQCR)
      { S7_Templates := "SrcType := Int" } GE_Contact(in1 := #STEP_30, in2 := #SQCR)
      Contact( "Clock_0.625Hz" )
   END_RUNG wire#w11
   RUNG wire#powerrail
      Contact( #smaz_me )
      Contact( "Clock_5Hz" )
      Coil( #smaz_me )
   END_RUNG
   RUNG wire#powerrail
      Contact( #smaz_me )
      Contact( "Clock_5Hz" )
      Coil( #smaz_me )
   END_RUNG
   // the same network as SCL:
   #_w1 := "alrm_global" OR "alrm_op_0" OR "alrm_op_1" OR "alrm_op_2" OR "alrm_op_3" OR "alrm_op_4" OR "alrm_op_5";
   #majak_red_s2 := #_w1 AND "Clock_1Hz";
   #majak_red_s3 := #majak_red_s2;
   #majak_red_s4 := #majak_red_s2;
   #majak_red_s5 := #majak_red_s2;
   #"M".hlaseni_chyby := #_w1;
   #"M".n_trig_wro := ("OP1_DB".TRIG.inicial_ok_op AND NOT #"M".hlaseni_chyby) OR ((#STEP_27 = #SQCR) AND "Clock_1Hz" AND "LOG_0") OR "DB_ALARM".ALARM.ALARM_GLOBAL OR ((#STEP_27 < #SQCR) AND "LOG_0") OR (("OP1_DB".SQCR > 5) AND ("OP1_DB".SQCR < 1000) AND "LOG_0") OR (("OP1_DB".SQCR = 5) AND ("OP1_DB".SQCR < 1000) AND "Clock_1Hz" AND "LOG_0");
   #majak_green_s1 := "AUTOMAT" AND (("OP1_DB".SQCR > 5) OR ("OP1_DB".SQCR = 5)) AND ("OP1_DB".SQCR < 1000);
   #majak_green_s2 := #majak_green_s1;
   #majak_green_s3 := #majak_green_s1;
   #majak_green_s4 := #majak_green_s1;
   #majak_green_s5 := #majak_green_s1;
   #"M".M_14 := "AUTOMAT" AND "alrm_global";
   #majak_blue_s1 := "AUTOMAT" AND ("OP1_DB".SQCR >= 1000) AND ("OP1_DB".SQCR <= 2000) AND NOT "DB_ALARM".ALARM.ALARM_GLOBAL;
   #majak_blue_s2 := #majak_blue_s1;
   #majak_blue_s3 := #majak_blue_s1;
   #majak_blue_s4 := #majak_blue_s1;
   #majak_blue_s5 := #majak_blue_s1;
   #majak_orange_s1 := "MANUAL";
   #majak_orange_s2 := "MANUAL";
   #majak_orange_s3 := "MANUAL";
   #majak_orange_s4 := "MANUAL";
   #majak_orange_s5 := "MANUAL";
   #majak_red_s1 := "AUTOMAT" AND "DB_ALARM".ALARM.ALARM_GLOBAL;
   #majak_red_s2 := #majak_red_s1;
   #majak_red_s3 := #majak_red_s1;
   #majak_red_s4 := #majak_red_s1;
   #majak_red_s5 := #majak_red_s1;
   #smaz_me := (#STEP_0_FIRST_START = #SQCR) OR ("DB_ALARM".ALARM.ALARM_GLOBAL AND "Clock_5Hz");
   #smaz_me := (#STEP_30 <= #SQCR) OR ((#STEP_0_FIRST_START <= #SQCR) AND (#STEP_30 >= #SQCR) AND "Clock_0.625Hz");
   #smaz_me := #smaz_me AND "Clock_5Hz";
   #smaz_me := #smaz_me AND "Clock_5Hz";
END_REGION

REGION Network 22: TRIG EXTERNAL
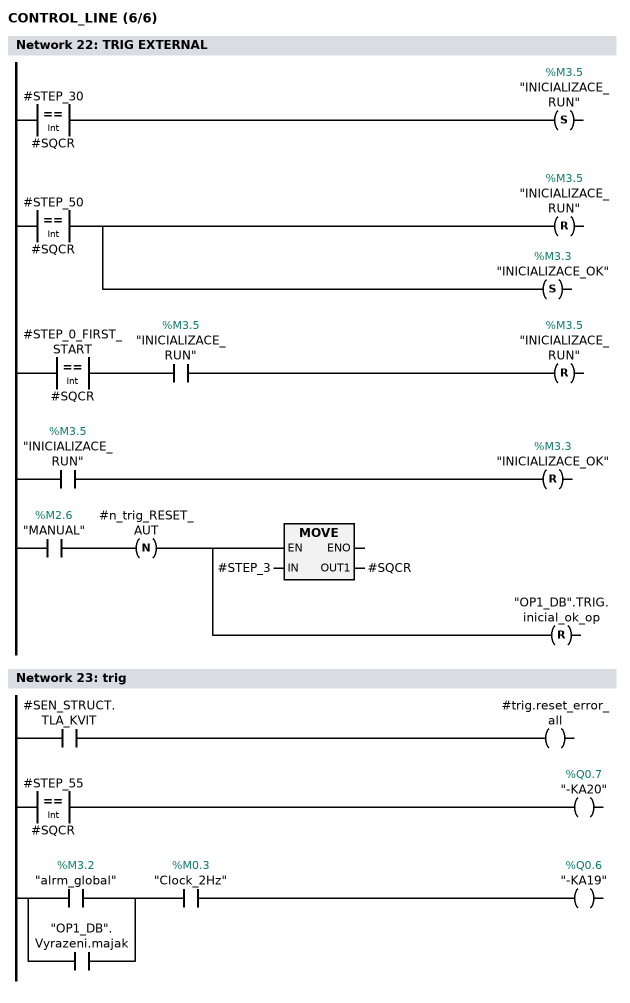
   RUNG wire#powerrail
      { S7_Templates := "SrcType := Int" } EQ_Contact(in1 := #STEP_30, in2 := #SQCR)
      S_Coil( "INICIALIZACE_RUN" )
   END_RUNG
   RUNG wire#powerrail
      { S7_Templates := "SrcType := Int" } EQ_Contact(in1 := #STEP_50, in2 := #SQCR)
      wire#w1
      R_Coil( "INICIALIZACE_RUN" )
   END_RUNG
   RUNG wire#w1
      S_Coil( "INICIALIZACE_OK" )
   END_RUNG
   RUNG wire#powerrail
      { S7_Templates := "SrcType := Int" } EQ_Contact(in1 := #STEP_0_FIRST_START, in2 := #SQCR)
      Contact( "INICIALIZACE_RUN" )
      R_Coil( "INICIALIZACE_RUN" )
   END_RUNG
   RUNG wire#powerrail
      Contact( "INICIALIZACE_RUN" )
      R_Coil( "INICIALIZACE_OK" )
   END_RUNG
   RUNG wire#powerrail
      Contact( "MANUAL" )
      N_Trig( #n_trig_RESET_AUT )
      wire#w2
      Move(in := #STEP_3, out1 => #SQCR)
   END_RUNG
   RUNG wire#w2
      R_Coil( "OP1_DB".TRIG.inicial_ok_op )
   END_RUNG
   // the same network as SCL:
   IF #STEP_30 = #SQCR THEN "INICIALIZACE_RUN" := TRUE; END_IF;
   IF #STEP_50 = #SQCR THEN
       "INICIALIZACE_RUN" := FALSE;
       "INICIALIZACE_OK" := TRUE;
   END_IF;
   IF (#STEP_0_FIRST_START = #SQCR) AND "INICIALIZACE_RUN" THEN "INICIALIZACE_RUN" := FALSE; END_IF;
   IF "INICIALIZACE_RUN" THEN "INICIALIZACE_OK" := FALSE; END_IF;
   #_w1 := NOT "MANUAL" AND #n_trig_RESET_AUT;   // falling edge
   #n_trig_RESET_AUT := "MANUAL";
   IF #_w1 THEN
       #SQCR := #STEP_3;
       "OP1_DB".TRIG.inicial_ok_op := FALSE;
   END_IF;
END_REGION

REGION Network 23: trig
   RUNG wire#powerrail
      Contact( #SEN_STRUCT.TLA_KVIT )
      Coil( #trig.reset_error_all )
   END_RUNG
   RUNG wire#powerrail
      { S7_Templates := "SrcType := Int" } EQ_Contact(in1 := #STEP_55, in2 := #SQCR)
      Coil( "-KA20" )
   END_RUNG
   RUNG wire#powerrail
      Contact( "alrm_global" )
      wire#w1
      Contact( "Clock_2Hz" )
      Coil( "-KA19" )
   END_RUNG
   RUNG wire#powerrail
      Contact( "OP1_DB".Vyrazeni.majak )
   END_RUNG wire#w1
   // the same network as SCL:
   #trig.reset_error_all := #SEN_STRUCT.TLA_KVIT;
   "-KA20" := #STEP_55 = #SQCR;
   "-KA19" := ("alrm_global" OR "OP1_DB".Vyrazeni.majak) AND "Clock_2Hz";
END_REGION
END_FUNCTION_BLOCK

FUNCTION_BLOCK "OP1"   // FB50, LAD
{ S7_Optimized_Access := 'TRUE' }
// stored: AutoNumber false, MemoryReserve 100, SetENOAutomatically false
   VAR DB_SPECIFIC
      CONTROL_MAN : Struct
         kar_work : Bool;
         kar_home : Bool;
         zarazka_work : Bool;
         zarazka_home : Bool;
         B4 : Bool;
         B5 : Bool;
         B6 : Bool;
         B7 : Bool;
         B8 : Bool;
         B9 : Bool;
         odfuk_1 : Bool;
         odfuk_2 : Bool;
         B12 : Bool;
         B13 : Bool;
         B14 : Bool;
         B15 : Bool;
         B16 : Bool;
         B17 : Bool;
         B18 : Bool;
         B19 : Bool;
         B20 : Bool;
         B21 : Bool;
         B22 : Bool;
         B23 : Bool;
         B24 : Bool;
         B25 : Bool;
         B26 : Bool;
         B27 : Bool;
         B28 : Bool;
         B29 : Bool;
         B30 : Bool;
         B31 : Bool;
      END_STRUCT;
      CONTROL_AUTOMAT : Struct
         KAR_WORK : Bool;
         KAR_HOME : Bool;
         ZARAZKA_WORK : Bool;
         ZARAZKA_HOME : Bool;
         B4 : Bool;
         B5 : Bool;
         B6 : Bool;
         B7 : Bool;
         B8 : Bool;
         B9 : Bool;
         odfuk_1 : Bool;
         odfuk_2 : Bool;
         B12 : Bool;
         B13 : Bool;
         B14 : Bool;
         B15 : Bool;
         B16 : Bool;
         B17 : Bool;
         B18 : Bool;
         B19 : Bool;
         B20 : Bool;
         B21 : Bool;
         B22 : Bool;
         B23 : Bool;
         B24 : Bool;
         B25 : Bool;
         B26 : Bool;
         B27 : Bool;
         B28 : Bool;
         B29 : Bool;
         B30 : Bool;
         B31 : Bool;
      END_STRUCT;
      SENSORS : Struct
         prechod_1 : Bool;
         prechod_1_neg : Bool;
         kontrola : Bool;
         kontrola_neg : Bool;
         prechod_2 : Bool;
         Prechod_2_neg : Bool;
         Pozice_vyrazovace : Bool;
         Pozice_vyrazovace_neg : Bool;
         Pozice_pistu : Bool;   // KARUSEL JE NATOČEN PŘÍPRAVKEM A K BRÁNĚ
         Pozice_pistu_neg : Bool;
         s10 : Bool;
         s11 : Bool;
         s12 : Bool;
         s13 : Bool;
         s14 : Bool;
         s15 : Bool;
         s16 : Bool;
         s17 : Bool;
         s18 : Bool;
         s19 : Bool;
         s20 : Bool;
         s21 : Bool;
         s22 : Bool;
         s23 : Bool;
         s24 : Bool;
         s25 : Bool;
         s26 : Bool;
         s27 : Bool;
         s28 : Bool;
         s29 : Bool;
         s30 : Bool;
         s31 : Bool;
      END_STRUCT;
      SENSORS_1 : Struct
         S0 : Bool;
         S1 : Bool;
         S2 : Bool;
         S3 : Bool;
         S4 : Bool;
         S5 : Bool;
         S6 : Bool;
         S7 : Bool;
         S8 : Bool;
         S9 : Bool;
         SESTAVA_NENI_OTOCENA : Bool;
         SESTAVA_JE_OTOCENA : Bool;
         S12 : Bool;
         S13 : Bool;
         S14 : Bool;
         S15 : Bool;
         S16 : Bool;
         S17 : Bool;
         S18 : Bool;
         S19 : Bool;
         S20 : Bool;
         S21 : Bool;
         S22 : Bool;
         S23 : Bool;
         S24 : Bool;
         S25 : Bool;
         S26 : Bool;
         S27 : Bool;
         S28 : Bool;
         S29 : Bool;
         S30 : Bool;
         l_3_neg : Bool;
      END_STRUCT;
   END_VAR
   VAR
      S_0 : "SENSOR";
      S_1 : "SENSOR";
      S_2 { S7_SetPoint := 'True'} : "SENSOR";
      S_3 { S7_SetPoint := 'True'} : "SENSOR";
      S_4 { S7_SetPoint := 'True'} : "SENSOR";
      S_5 { S7_SetPoint := 'True'} : "SENSOR";
      S_6 { S7_SetPoint := 'True'} : "SENSOR";
      M_karusel : "MOTOR_CONTROL_BLOCK";
      M_zarazka { S7_SetPoint := 'True'} : "MOTOR_CONTROL_BLOCK";
      M_CLONA { S7_SetPoint := 'True'} : "MOTOR_CONTROL_BLOCK";
   END_VAR
   VAR DB_SPECIFIC
      SQCR { S7_SetPoint := 'True'} : Int;
   END_VAR
   VAR
      hmi_sqcr : Int;
   END_VAR
   VAR DB_SPECIFIC
      TRIG : Struct
         inicial_ok_op : Bool;
         DSSAD : Bool;
         INICIALIZACE_PROBEHLA : Bool;
         trig_dil : Bool;
         p_trig_control_tcon : Bool;
         T6 : Bool;
         SPUST_OP_4 : Bool;
         vlez_do_zavory_pri_rotaci : Bool;
         START_INICIAL_OP2 : Bool;
         START_INICIAL_OP3 : Bool;
         spust_odsavani : Bool;
         VYPRAZNI_OK_OP_2_A : Bool;
         VYPRAZNI_NOK_OP_2_A : Bool;
         VYPRAZDNI_OK_OP_3_B : Bool;
         VYPRAZDNI_NOK_OP_3_B : Bool;
         RESET_NCODER : Bool;
         op_1_ready : Bool;
      END_STRUCT;
      MEMOR : Struct
         n_trig_vypnuti : Bool;
         M1 : Bool;
         M2 : Bool;
         M3 : Bool;
         M4 : Bool;
         p_trig_odavacka : Bool;
         M6 : Bool;
         M7 : Bool;
         M8 : Bool;
         M9 : Bool;
         M10 : Bool;
         M11 : Bool;
         RESET_ERROR : Bool;
         vyrazeni_pamet : Bool;
         M14 : Bool;
         M15 : Bool;
         SETOVANI_START : Bool;
         M17 : Bool;
         p_trig_pamet_1 : Bool;
         p_trig_pamet_2 : Bool;
         p_trig_pamet_3 : Bool;
         p_trig_pamet_4 : Bool;
         p_trig_pamet_5 : Bool;
         p_trig_pamet_6 : Bool;
         p_trig_pamet_7 : Bool;
         p_trig_pamet_8 : Bool;
         p_trig_pamet_9 : Bool;
         p_trig_pamet_10 : Bool;
         p_trig_vyrad : Bool;
         p_Trig_cisteni_pozice : Bool;
         p_trig_citac : Bool;
         N_TRIG_SAFETY : Bool;
         P_TRIG_RESET_POZICE : Bool;
         M33 : Bool;
         start_caklu : Bool;
         M35 : Bool;
         M36 : Bool;
         M37 : Bool;
         M38 : Bool;
         M39 : Bool;
         ALARM_GLOBAL : Bool;
         M41 : Bool;
         M42 : Bool;
         M43 : Bool;
         M44 : Bool;
         M45 : Bool;
         M46 : Bool;
         M47 : Bool;
         M48 : Bool;
         M49 : Bool;
         wrong_p_trig : Bool;
         alarm_p_trig : Bool;
         M52 : Bool;
         M53 : Bool;
         M54 : Bool;
         M55 : Bool;
         M56 : Bool;
         M57 : Bool;
         M58 : Bool;
         M59 : Bool;
         M60 : Bool;
         M61 : Bool;
         M62 : Bool;
         M63 : Bool;
      END_STRUCT;
      "TIMER" : Struct
         TIMER_0 : IEC_TIMER;
         TIMER_VACUUM_CLEANER : IEC_TIMER;
         TIMER_DELAY_RESET_EXECUTE : IEC_TIMER;
         TIMER_3 : IEC_TIMER;
         TIMER_4 : IEC_TIMER;
         air : IEC_TIMER;
         TIMER_6 : IEC_TIMER;
         TIMER_7 : IEC_TIMER;
      END_STRUCT;
      HMI : Struct
         povoleni_volby_receptu : Bool;
         "svetlo_on/off" : Bool;
         ALARM_VIDITELNOST : Bool;
         hmi_3 : Bool;
         hmi_4 : Bool;
         reset_fronty : Bool;
         hmi_6 : Bool;
         hmi_7 : Bool;
         hmi_8 : Bool;
         hmi_9 : Bool;
         hmi_10 : Bool;
         hmi_11 : Bool;
         hmi_12 : Bool;
         hmi_13 : Bool;
         hmi_14 : Bool;
         hmi_15 : Bool;
      END_STRUCT;
   END_VAR
   VAR
      STRING_0 : String[1];
      array_chyb_ctec : Array[1..16] of Bool;
      zpracovani_dat { ExternalAccessible := 'False'; ExternalVisible := 'False'; ExternalWritable := 'False'} : Array[1..1] of Struct
         prenaseny_text : String[100];
         balik_den : Int;
         vyrazeni : Bool;
      END_STRUCT;
   END_VAR
   VAR DB_SPECIFIC
      aktual_kusy : Int;
   END_VAR
   VAR
      i : Int;
      q : Int;
      pocet_znaku_string_kamera : Int;
      ocekavany_text : String[100];
      format_etiketa_ok : Bool;
      Kamera : Struct
         s2_pamet : Bool;
         s2_nabeh : Bool;
         sber_aktivni : Bool;
         prijato_etiketa : Bool;
         prijato_folie_l : Bool;
         prijato_folie_p : Bool;
         ok_etiketa : Bool;
         ok_folie_l : Bool;
         ok_folie_p : Bool;
         vyradit : Bool;
         fronta_plna : Bool;   // alarm
         bypass_ocr : Bool := True;   // dočasně, dokud není doladěné OCR
         last_id_etiketa : Word;
         last_id_folie_l : Word;
         last_id_folie_p : Word;
         balik_den : Int;
         idx : Int;
         pocet : Int;
         text_etiketa : String[100];
         timeout_sberu : Time :=  T#1S;
         kontrola_tridirny : Bool := true;   // HMI: kontrola kódu třídírny zapnuta
         tridirna_ok : Bool;   // výsledek kontroly posledního plata (pro online diagnostiku)
      END_STRUCT;
      Vyrazeni : Struct
         s4_pamet : Bool;
         s4_nabeh : Bool;
         aktivni : Bool;
         vyradit : Bool;
         chyba_bez_dat : Bool;   // alarm: plato u vyřazovače bez záznamu
         chyba_pist : Bool;   // alarm: píst nevyjel / nebyl v home
         max_puls : Time := T#200MS;
         vyrazovac_pripojen : Bool := true;   // TRUE až bude signál od dodavatele
         alarm_nok_balik : Bool;   // NOK plato prošlo bez vyřazení
         posledni_nok_balik : Int;   // číslo plata pro obsluhu / HMI
         posledni_nok_text : String[100];   // co přečetla kamera
         pocet_nok : DInt;   // počítadlo NOK plat
         pocet_bez_dat : DInt;
         majak_tp : TP_TIME;   // prodlouzeni blikani majaku pri vzrazenii
         majak { S7_SetPoint := 'True'} : Bool;
      END_STRUCT;
      Kam_Etiketa_Job : Struct
         krok : Int;   // 0 klid, 10 odeslat, 20 čekat, 30 ukončit handshake
         pozadovany : Int;   // job z receptury (PRG_CAM_etiketa)
         odesli_pamet : Bool;   // hrana ODESLI_dATA
         aktivni : Bool;   // probíhá načítání jobu → blokovat triggery
         chyba : Bool;   // alarm: job se nepodařilo načíst
         chyba_kod : Word;   // CommandResultCode při chybě
         nesouhlasi : Bool;   // alarm: job v kameře ≠ job z receptury
         timeout : Time := T#10S;   // max. doba načítání jobu
      END_STRUCT;
      Test_tp_ka12 : TP_TIME;
   END_VAR
   VAR_TEMP
      DATA : Array[0..255] of Char;
      ARRAY_NULL : Array[1..8] of Bool;
      array_null_fronta : Array[1..1] of Struct
         prenaseny_text : String[100];
         balik_den : Int;
         vyrazeni : Bool;
      END_STRUCT;
      "char" : Array[0..0] of Char;
      "string" : String;
      cas : DTL;
      ret : Int;
   END_VAR
   VAR CONSTANT
      STEP_0 : Int := 0;
      step_2 : Int := 2;
      STEP_4 : Int := 4;
      STEP_5_HOME : Int := 5;
      STEP_7 : Int := 7;
      STEP_10 : Int := 10;
      STEP_15 : Int := 15;
      STEP_20 : Int := 20;
      STEP_23 : Int := 23;
      STEP_25 : Int := 25;
      STEP_27 : Int := 27;
      STEP_30 : Int := 30;
      STEP_35 : Int := 35;
      STEP_37 : Int := 37;
      STEP_40 : Int := 40;
      STEP_45 : Int := 45;
      STEP_50 : Int := 50;
      STEP_55 : Int := 55;
      STEP_60 : Int := 60;
      STEP_65 : Int := 65;
      STEP_70 : Int := 70;
      STEP_75 : Int := 75;
      STEP_80 : Int := 80;
      STEP_83 : Int := 83;
      STEP_85 : Int := 85;
      STEP_90 : Int := 90;
      STEP_95 : Int := 95;
      STEP_100 : Int := 100;
      STEP_105 : Int := 105;
      STEP_110 : Int := 110;
      STEP_113 : Int := 113;
      STEP_115 : Int := 115;
      STEP_120 : Int := 120;
      STEP_125 : Int := 125;
      STEP_130 : Int := 130;
      STEP_135 : Int := 135;
      STEP_140 : Int := 140;
      STEP_145 : Int := 145;
      STEP_150 : Int := 150;
      STEP_155 : Int := 155;
      STEP_1000 : Int := 1000;
      STEP_1001 : Int := 1001;
      STEP_1002 : Int := 1002;
      STEP_1003 : Int := 1003;
      STEP_1004 : Int := 1004;
      STEP_1005 : Int := 1005;
      STEP_1010 : Int := 1010;
      STEP_1015 : Int := 1015;
      STEP_1020 : Int := 1020;
      STEP_1025 : Int := 1025;
      STEP_3000 : Int := 3000;
      STEP_3005 : Int := 3005;
      STEP_3010 : Int := 3010;
      STEP_3015 : Int := 3015;
      STEP_3020 : Int := 3020;
      STEP_2000 : Int := 2000;
      string_null : String;
      char_null : Char;
      text_kartacek : String := 'Kartacek';
      string_kar_A : String := 'A';
      string_kar_B : String := 'B';
      KOD_TRIDIRNY : String := 'CZ32880102';
   END_VAR
   VAR_TEMP   // added for the SCL form of the ladder/FBD networks
      _w1 : Bool;
      _w2 : Bool;
      _w3 : Bool;
   END_VAR
BEGIN

REGION Network 1: manuali ovladani reset
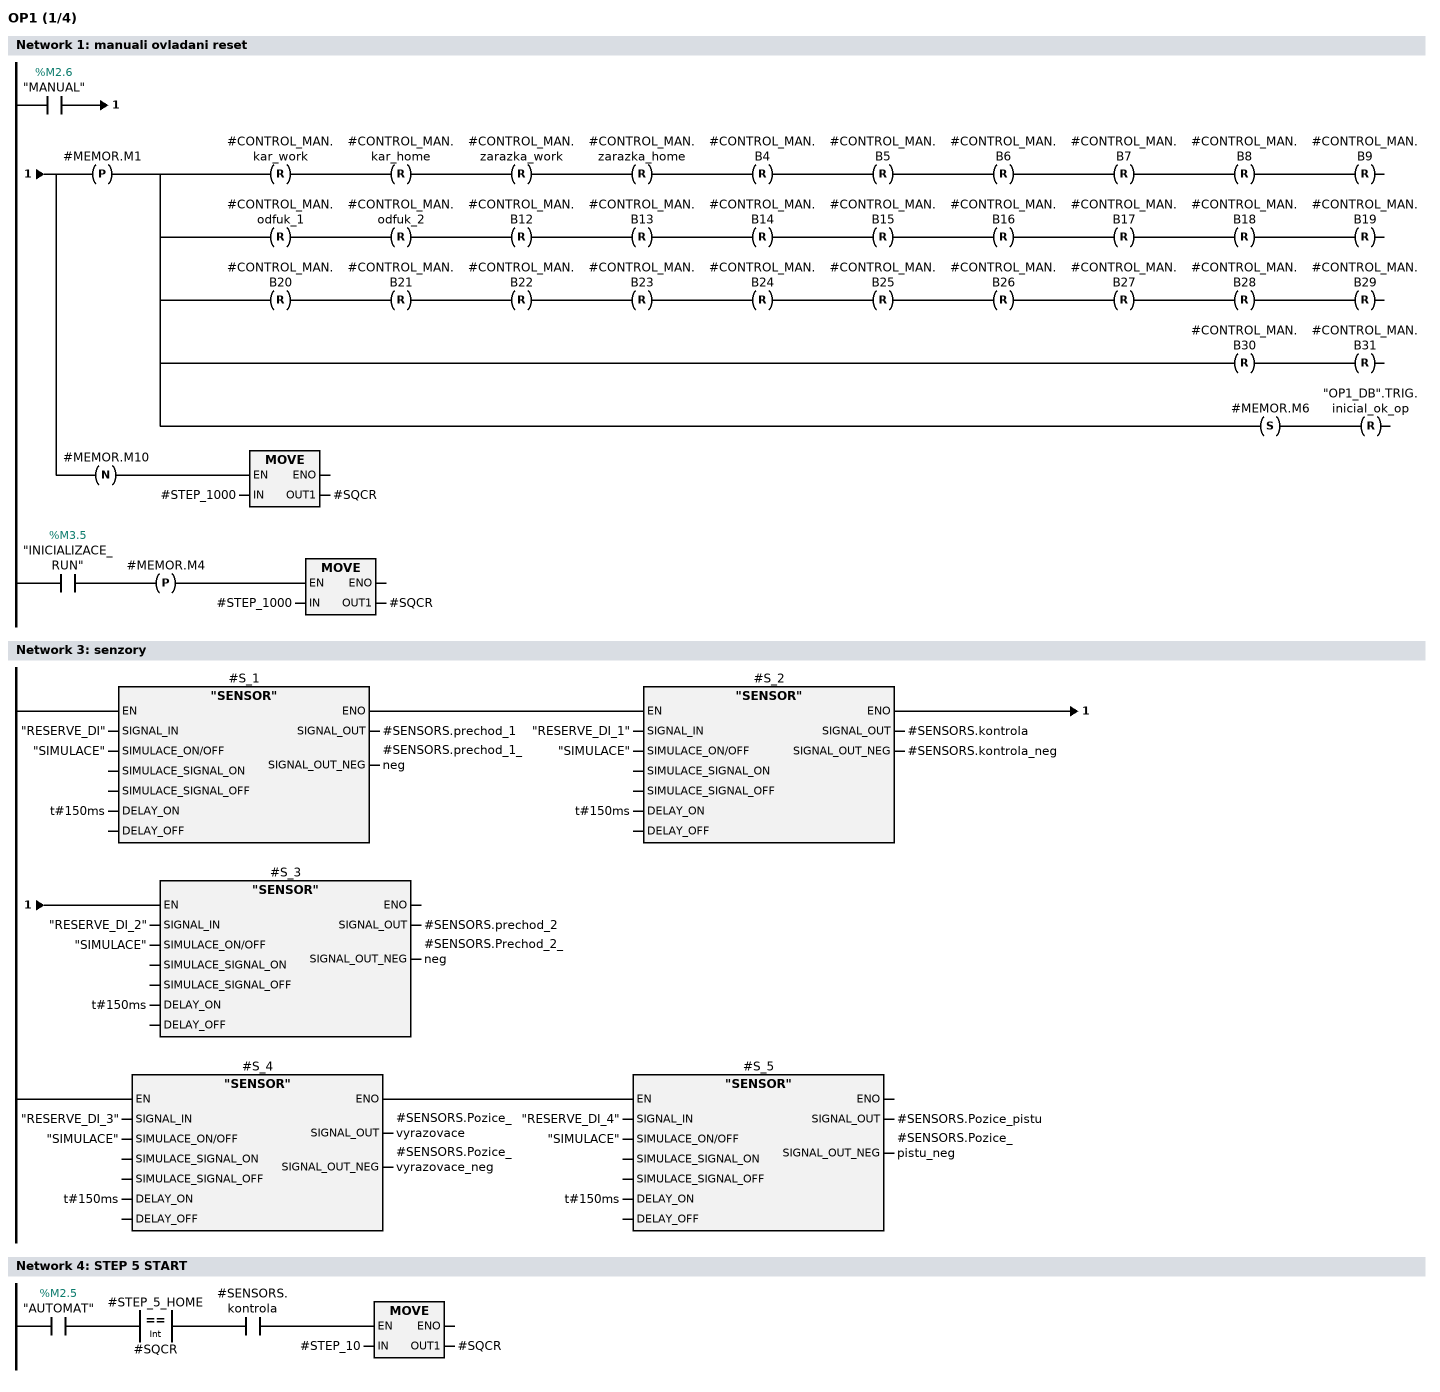
   RUNG wire#powerrail
      Contact( "MANUAL" )
      wire#w1
      P_Trig( #MEMOR.M1 )
      wire#w2
      R_Coil( #CONTROL_MAN.kar_work )
      R_Coil( #CONTROL_MAN.kar_home )
      R_Coil( #CONTROL_MAN.zarazka_work )
      R_Coil( #CONTROL_MAN.zarazka_home )
      R_Coil( #CONTROL_MAN.B4 )
      R_Coil( #CONTROL_MAN.B5 )
      R_Coil( #CONTROL_MAN.B6 )
      R_Coil( #CONTROL_MAN.B7 )
      R_Coil( #CONTROL_MAN.B8 )
      R_Coil( #CONTROL_MAN.B9 )
   END_RUNG
   RUNG wire#w2
      R_Coil( #CONTROL_MAN.odfuk_1 )
      R_Coil( #CONTROL_MAN.odfuk_2 )
      R_Coil( #CONTROL_MAN.B12 )
      R_Coil( #CONTROL_MAN.B13 )
      R_Coil( #CONTROL_MAN.B14 )
      R_Coil( #CONTROL_MAN.B15 )
      R_Coil( #CONTROL_MAN.B16 )
      R_Coil( #CONTROL_MAN.B17 )
      R_Coil( #CONTROL_MAN.B18 )
      R_Coil( #CONTROL_MAN.B19 )
   END_RUNG
   RUNG wire#w2
      R_Coil( #CONTROL_MAN.B20 )
      R_Coil( #CONTROL_MAN.B21 )
      R_Coil( #CONTROL_MAN.B22 )
      R_Coil( #CONTROL_MAN.B23 )
      R_Coil( #CONTROL_MAN.B24 )
      R_Coil( #CONTROL_MAN.B25 )
      R_Coil( #CONTROL_MAN.B26 )
      R_Coil( #CONTROL_MAN.B27 )
      R_Coil( #CONTROL_MAN.B28 )
      R_Coil( #CONTROL_MAN.B29 )
   END_RUNG
   RUNG wire#w2
      R_Coil( #CONTROL_MAN.B30 )
      R_Coil( #CONTROL_MAN.B31 )
   END_RUNG
   RUNG wire#w2
      S_Coil( #MEMOR.M6 )
      R_Coil( "OP1_DB".TRIG.inicial_ok_op )
   END_RUNG
   RUNG wire#w1
      N_Trig( #MEMOR.M10 )
      Move(in := #STEP_1000, out1 => #SQCR)
   END_RUNG
   RUNG wire#powerrail
      Contact( "INICIALIZACE_RUN" )
      P_Trig( #MEMOR.M4 )
      Move(in := #STEP_1000, out1 => #SQCR)
   END_RUNG
   // the same network as SCL:
   #_w1 := "MANUAL" AND NOT #MEMOR.M1;   // rising edge
   #MEMOR.M1 := "MANUAL";
   IF #_w1 THEN
       #CONTROL_MAN.kar_work := FALSE;
       #CONTROL_MAN.kar_home := FALSE;
       #CONTROL_MAN.zarazka_work := FALSE;
       #CONTROL_MAN.zarazka_home := FALSE;
       #CONTROL_MAN.B4 := FALSE;
       #CONTROL_MAN.B5 := FALSE;
       #CONTROL_MAN.B6 := FALSE;
       #CONTROL_MAN.B7 := FALSE;
       #CONTROL_MAN.B8 := FALSE;
       #CONTROL_MAN.B9 := FALSE;
       #CONTROL_MAN.odfuk_1 := FALSE;
       #CONTROL_MAN.odfuk_2 := FALSE;
       #CONTROL_MAN.B12 := FALSE;
       #CONTROL_MAN.B13 := FALSE;
       #CONTROL_MAN.B14 := FALSE;
       #CONTROL_MAN.B15 := FALSE;
       #CONTROL_MAN.B16 := FALSE;
       #CONTROL_MAN.B17 := FALSE;
       #CONTROL_MAN.B18 := FALSE;
       #CONTROL_MAN.B19 := FALSE;
       #CONTROL_MAN.B20 := FALSE;
       #CONTROL_MAN.B21 := FALSE;
       #CONTROL_MAN.B22 := FALSE;
       #CONTROL_MAN.B23 := FALSE;
       #CONTROL_MAN.B24 := FALSE;
       #CONTROL_MAN.B25 := FALSE;
       #CONTROL_MAN.B26 := FALSE;
       #CONTROL_MAN.B27 := FALSE;
       #CONTROL_MAN.B28 := FALSE;
       #CONTROL_MAN.B29 := FALSE;
       #CONTROL_MAN.B30 := FALSE;
       #CONTROL_MAN.B31 := FALSE;
       #MEMOR.M6 := TRUE;
       "OP1_DB".TRIG.inicial_ok_op := FALSE;
   END_IF;
   #_w2 := NOT "MANUAL" AND #MEMOR.M10;   // falling edge
   #MEMOR.M10 := "MANUAL";
   IF #_w2 THEN #SQCR := #STEP_1000; END_IF;
   #_w3 := "INICIALIZACE_RUN" AND NOT #MEMOR.M4;   // rising edge
   #MEMOR.M4 := "INICIALIZACE_RUN";
   IF #_w3 THEN #SQCR := #STEP_1000; END_IF;
END_REGION

REGION Network 2: alarmy
END_REGION

REGION Network 3: senzory
   RUNG wire#powerrail
      #S_1(SIGNAL_IN := "RESERVE_DI", "SIMULACE_ON/OFF" := "SIMULACE", SIMULACE_SIGNAL_ON :=, SIMULACE_SIGNAL_OFF :=, DELAY_ON := t#150ms, DELAY_OFF :=, SIGNAL_OUT => #SENSORS.prechod_1, SIGNAL_OUT_NEG => #SENSORS.prechod_1_neg)
      #S_2(SIGNAL_IN := "RESERVE_DI_1", "SIMULACE_ON/OFF" := "SIMULACE", SIMULACE_SIGNAL_ON :=, SIMULACE_SIGNAL_OFF :=, DELAY_ON := t#150ms, DELAY_OFF :=, SIGNAL_OUT => #SENSORS.kontrola, SIGNAL_OUT_NEG => #SENSORS.kontrola_neg)
      #S_3(SIGNAL_IN := "RESERVE_DI_2", "SIMULACE_ON/OFF" := "SIMULACE", SIMULACE_SIGNAL_ON :=, SIMULACE_SIGNAL_OFF :=, DELAY_ON := t#150ms, DELAY_OFF :=, SIGNAL_OUT => #SENSORS.prechod_2, SIGNAL_OUT_NEG => #SENSORS.Prechod_2_neg)
   END_RUNG
   RUNG wire#powerrail
      #S_4(SIGNAL_IN := "RESERVE_DI_3", "SIMULACE_ON/OFF" := "SIMULACE", SIMULACE_SIGNAL_ON :=, SIMULACE_SIGNAL_OFF :=, DELAY_ON := t#150ms, DELAY_OFF :=, SIGNAL_OUT => #SENSORS.Pozice_vyrazovace, SIGNAL_OUT_NEG => #SENSORS.Pozice_vyrazovace_neg)
      #S_5(SIGNAL_IN := "RESERVE_DI_4", "SIMULACE_ON/OFF" := "SIMULACE", SIMULACE_SIGNAL_ON :=, SIMULACE_SIGNAL_OFF :=, DELAY_ON := t#150ms, DELAY_OFF :=, SIGNAL_OUT => #SENSORS.Pozice_pistu, SIGNAL_OUT_NEG => #SENSORS.Pozice_pistu_neg)
   END_RUNG
   // the same network as SCL:
   #S_1(SIGNAL_IN := "RESERVE_DI",   // "SENSOR"
        "SIMULACE_ON/OFF" := "SIMULACE",
        DELAY_ON := t#150ms,
        SIGNAL_OUT => #SENSORS.prechod_1,
        SIGNAL_OUT_NEG => #SENSORS.prechod_1_neg,
        ENO => #_w1);
   #S_2(EN := #_w1,   // "SENSOR"
        SIGNAL_IN := "RESERVE_DI_1",
        "SIMULACE_ON/OFF" := "SIMULACE",
        DELAY_ON := t#150ms,
        SIGNAL_OUT => #SENSORS.kontrola,
        SIGNAL_OUT_NEG => #SENSORS.kontrola_neg,
        ENO => #_w2);
   IF #_w2 THEN
       #S_3(SIGNAL_IN := "RESERVE_DI_2",   // "SENSOR"
            "SIMULACE_ON/OFF" := "SIMULACE",
            DELAY_ON := t#150ms,
            SIGNAL_OUT => #SENSORS.prechod_2,
            SIGNAL_OUT_NEG => #SENSORS.Prechod_2_neg);
   END_IF;
   #S_4(SIGNAL_IN := "RESERVE_DI_3",   // "SENSOR"
        "SIMULACE_ON/OFF" := "SIMULACE",
        DELAY_ON := t#150ms,
        SIGNAL_OUT => #SENSORS.Pozice_vyrazovace,
        SIGNAL_OUT_NEG => #SENSORS.Pozice_vyrazovace_neg,
        ENO => #_w3);
   IF #_w3 THEN
       #S_5(SIGNAL_IN := "RESERVE_DI_4",   // "SENSOR"
            "SIMULACE_ON/OFF" := "SIMULACE",
            DELAY_ON := t#150ms,
            SIGNAL_OUT => #SENSORS.Pozice_pistu,
            SIGNAL_OUT_NEG => #SENSORS.Pozice_pistu_neg);
   END_IF;
END_REGION

REGION Network 4: STEP 5 START
   RUNG wire#powerrail
      Contact( "AUTOMAT" )
      { S7_Templates := "SrcType := Int" } EQ_Contact(in1 := #STEP_5_HOME, in2 := #SQCR)
      Contact( #SENSORS.kontrola )
      Move(in := #STEP_10, out1 => #SQCR)
   END_RUNG
   // the same network as SCL:
   IF "AUTOMAT" AND (#STEP_5_HOME = #SQCR) AND #SENSORS.kontrola THEN #SQCR := #STEP_10; END_IF;
END_REGION

REGION Network 5: STEP 10
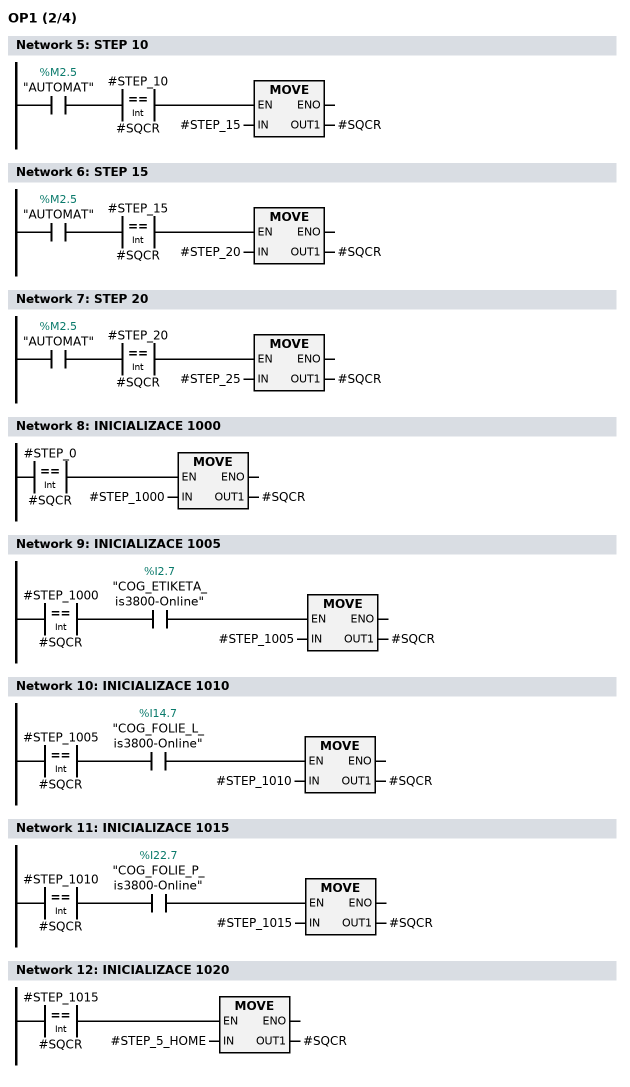
   RUNG wire#powerrail
      Contact( "AUTOMAT" )
      { S7_Templates := "SrcType := Int" } EQ_Contact(in1 := #STEP_10, in2 := #SQCR)
      Move(in := #STEP_15, out1 => #SQCR)
   END_RUNG
   // the same network as SCL:
   IF "AUTOMAT" AND (#STEP_10 = #SQCR) THEN #SQCR := #STEP_15; END_IF;
END_REGION

REGION Network 6: STEP 15
   RUNG wire#powerrail
      Contact( "AUTOMAT" )
      { S7_Templates := "SrcType := Int" } EQ_Contact(in1 := #STEP_15, in2 := #SQCR)
      Move(in := #STEP_20, out1 => #SQCR)
   END_RUNG
   // the same network as SCL:
   IF "AUTOMAT" AND (#STEP_15 = #SQCR) THEN #SQCR := #STEP_20; END_IF;
END_REGION

REGION Network 7: STEP 20
   RUNG wire#powerrail
      Contact( "AUTOMAT" )
      { S7_Templates := "SrcType := Int" } EQ_Contact(in1 := #STEP_20, in2 := #SQCR)
      Move(in := #STEP_25, out1 => #SQCR)
   END_RUNG
   // the same network as SCL:
   IF "AUTOMAT" AND (#STEP_20 = #SQCR) THEN #SQCR := #STEP_25; END_IF;
END_REGION

REGION Network 8: INICIALIZACE 1000
   RUNG wire#powerrail
      { S7_Templates := "SrcType := Int" } EQ_Contact(in1 := #STEP_0, in2 := #SQCR)
      Move(in := #STEP_1000, out1 => #SQCR)
   END_RUNG
   // the same network as SCL:
   IF #STEP_0 = #SQCR THEN #SQCR := #STEP_1000; END_IF;
END_REGION

REGION Network 9: INICIALIZACE 1005
   RUNG wire#powerrail
      { S7_Templates := "SrcType := Int" } EQ_Contact(in1 := #STEP_1000, in2 := #SQCR)
      Contact( "COG_ETIKETA_is3800-Online" )
      Move(in := #STEP_1005, out1 => #SQCR)
   END_RUNG
   // the same network as SCL:
   IF (#STEP_1000 = #SQCR) AND "COG_ETIKETA_is3800-Online" THEN #SQCR := #STEP_1005; END_IF;
END_REGION

REGION Network 10: INICIALIZACE 1010
   RUNG wire#powerrail
      { S7_Templates := "SrcType := Int" } EQ_Contact(in1 := #STEP_1005, in2 := #SQCR)
      Contact( "COG_FOLIE_L_is3800-Online" )
      Move(in := #STEP_1010, out1 => #SQCR)
   END_RUNG
   // the same network as SCL:
   IF (#STEP_1005 = #SQCR) AND "COG_FOLIE_L_is3800-Online" THEN #SQCR := #STEP_1010; END_IF;
END_REGION

REGION Network 11: INICIALIZACE 1015
   RUNG wire#powerrail
      { S7_Templates := "SrcType := Int" } EQ_Contact(in1 := #STEP_1010, in2 := #SQCR)
      Contact( "COG_FOLIE_P_is3800-Online" )
      Move(in := #STEP_1015, out1 => #SQCR)
   END_RUNG
   // the same network as SCL:
   IF (#STEP_1010 = #SQCR) AND "COG_FOLIE_P_is3800-Online" THEN #SQCR := #STEP_1015; END_IF;
END_REGION

REGION Network 12: INICIALIZACE 1020
   RUNG wire#powerrail
      { S7_Templates := "SrcType := Int" } EQ_Contact(in1 := #STEP_1015, in2 := #SQCR)
      Move(in := #STEP_5_HOME, out1 => #SQCR)
   END_RUNG
   // the same network as SCL:
   IF #STEP_1015 = #SQCR THEN #SQCR := #STEP_5_HOME; END_IF;
END_REGION

REGION Network 13: automat control door / TRIGGER KAMER
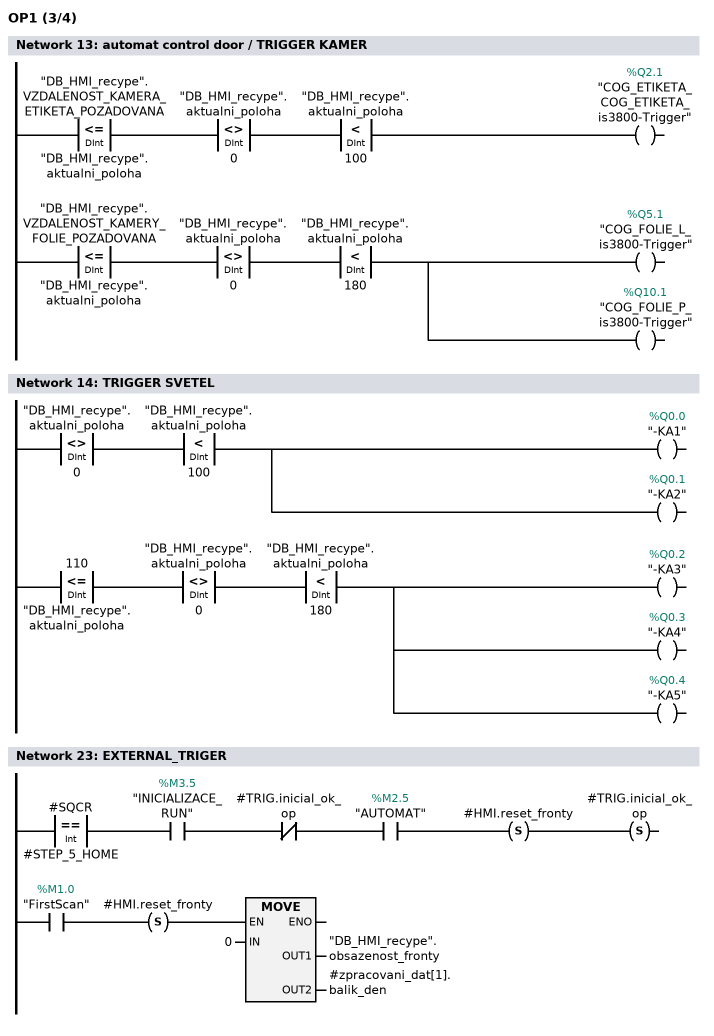
   RUNG wire#powerrail
      { S7_Templates := "SrcType := DInt" } LE_Contact(in1 := "DB_HMI_recype".VZDALENOST_KAMERA_ETIKETA_POZADOVANA, in2 := "DB_HMI_recype".aktualni_poloha)
      { S7_Templates := "SrcType := DInt" } NE_Contact(in1 := "DB_HMI_recype".aktualni_poloha, in2 := 0)
      { S7_Templates := "SrcType := DInt" } LT_Contact(in1 := "DB_HMI_recype".aktualni_poloha, in2 := 100)
      Coil( "COG_ETIKETA_COG_ETIKETA_is3800-Trigger" )
   END_RUNG
   RUNG wire#powerrail
      { S7_Templates := "SrcType := DInt" } LE_Contact(in1 := "DB_HMI_recype".VZDALENOST_KAMERY_FOLIE_POZADOVANA, in2 := "DB_HMI_recype".aktualni_poloha)
      { S7_Templates := "SrcType := DInt" } NE_Contact(in1 := "DB_HMI_recype".aktualni_poloha, in2 := 0)
      { S7_Templates := "SrcType := DInt" } LT_Contact(in1 := "DB_HMI_recype".aktualni_poloha, in2 := 180)
      wire#w1
      Coil( "COG_FOLIE_L_is3800-Trigger" )
   END_RUNG
   RUNG wire#w1
      Coil( "COG_FOLIE_P_is3800-Trigger" )
   END_RUNG
   // the same network as SCL:
   "COG_ETIKETA_COG_ETIKETA_is3800-Trigger" := ("DB_HMI_recype".VZDALENOST_KAMERA_ETIKETA_POZADOVANA <= "DB_HMI_recype".aktualni_poloha) AND ("DB_HMI_recype".aktualni_poloha <> 0) AND ("DB_HMI_recype".aktualni_poloha < 100);
   "COG_FOLIE_L_is3800-Trigger" := ("DB_HMI_recype".VZDALENOST_KAMERY_FOLIE_POZADOVANA <= "DB_HMI_recype".aktualni_poloha) AND ("DB_HMI_recype".aktualni_poloha <> 0) AND ("DB_HMI_recype".aktualni_poloha < 180);
   "COG_FOLIE_P_is3800-Trigger" := "COG_FOLIE_L_is3800-Trigger";
END_REGION

REGION Network 14: TRIGGER SVETEL
   RUNG wire#powerrail
      { S7_Templates := "SrcType := DInt" } NE_Contact(in1 := "DB_HMI_recype".aktualni_poloha, in2 := 0)
      { S7_Templates := "SrcType := DInt" } LT_Contact(in1 := "DB_HMI_recype".aktualni_poloha, in2 := 100)
      wire#w1
      Coil( "-KA1" )
   END_RUNG
   RUNG wire#w1
      Coil( "-KA2" )
   END_RUNG
   RUNG wire#powerrail
      { S7_Templates := "SrcType := DInt" } LE_Contact(in1 := 110, in2 := "DB_HMI_recype".aktualni_poloha)
      { S7_Templates := "SrcType := DInt" } NE_Contact(in1 := "DB_HMI_recype".aktualni_poloha, in2 := 0)
      { S7_Templates := "SrcType := DInt" } LT_Contact(in1 := "DB_HMI_recype".aktualni_poloha, in2 := 180)
      wire#w2
      Coil( "-KA3" )
   END_RUNG
   RUNG wire#w2
      Coil( "-KA4" )
   END_RUNG
   RUNG wire#w2
      Coil( "-KA5" )
   END_RUNG
   // the same network as SCL:
   "-KA1" := ("DB_HMI_recype".aktualni_poloha <> 0) AND ("DB_HMI_recype".aktualni_poloha < 100);
   "-KA2" := "-KA1";
   "-KA3" := (110 <= "DB_HMI_recype".aktualni_poloha) AND ("DB_HMI_recype".aktualni_poloha <> 0) AND ("DB_HMI_recype".aktualni_poloha < 180);
   "-KA4" := "-KA3";
   "-KA5" := "-KA3";
END_REGION

REGION Network 15 (SCL): TRIGGER MANUAL
   "iDB_CamManual"(xManEtiketa:="DB_Manual".xManEtiketa,
                   xManFolie:="DB_Manual".xManFolie);
END_REGION

REGION Network 16 (SCL): automat control data
   // Smyčka projde 104 bajtů (od 0 do 103)
   FOR #i := 0 TO 103 DO
       // PEEK čte přímo z paměti vstupů (16#81 = Periferní vstupy / Vstupy)
       // area 16#81 čte adresy %IB
       "DB_data_ctena".array_of_char[#i] := PEEK_BYTE(area := 16#81,
                                                       dbNumber := 0,
                                                       byteOffset := 76 + #i);
   END_FOR;

   // slozit text z prijatych znaku az po prvni $00
   "DB_data_ctena".upraveny := '';
   FOR #i := 0 TO 103 DO
       IF "DB_data_ctena".array_of_char[#i] = '$00' THEN
           EXIT;
       END_IF;
       "DB_data_ctena".upraveny := CONCAT(IN1 := "DB_data_ctena".upraveny,
                                          IN2 := CHAR_TO_STRING("DB_data_ctena".array_of_char[#i]));
   END_FOR;
END_REGION

REGION Network 17: automat control odfuk
END_REGION

REGION Network 18 (SCL): VYŘAZENÍ
   #Vyrazeni.s4_nabeh := #SENSORS.Pozice_vyrazovace AND NOT #Vyrazeni.s4_pamet;
   #Vyrazeni.s4_pamet := #SENSORS.Pozice_vyrazovace;

   IF "CONTROL_LINE_DB".trig.reset_error_all THEN
       #Vyrazeni.chyba_bez_dat := FALSE;
       #Vyrazeni.chyba_pist := FALSE;
       #Vyrazeni.alarm_nok_balik := FALSE;
   END_IF;

   IF NOT "AUTOMAT" THEN
       #Vyrazeni.aktivni := FALSE;
       #TIMER.TIMER_7.TON(IN := FALSE,
                          PT := #Vyrazeni.max_puls);
   ELSE
       REGION Plato prijelo k vyrazovaci - vzdy spotrebovat fronta[1]
           IF #Vyrazeni.s4_nabeh THEN
               IF "DB_HMI_recype".fronta[1].prenaseny_text = '' THEN
                   #Vyrazeni.chyba_bez_dat := TRUE;    // plato bez zaznamu ve fronte
                   #Vyrazeni.pocet_bez_dat := #Vyrazeni.pocet_bez_dat + 1;
                   #Vyrazeni.vyradit := TRUE;
               ELSE
                   #Vyrazeni.vyradit := "DB_HMI_recype".fronta[1].vyrazeni;
               END_IF;

               IF #Vyrazeni.vyradit THEN
                   #Vyrazeni.pocet_nok := #Vyrazeni.pocet_nok + 1;
                   IF "DB_HMI_recype".fronta[1].prenaseny_text = '' THEN
                       #Vyrazeni.posledni_nok_text := 'BEZ ZAZNAMU';
                       #Vyrazeni.posledni_nok_balik := 0;
                   ELSE
                       #Vyrazeni.posledni_nok_text := "DB_HMI_recype".fronta[1].prenaseny_text;
                       #Vyrazeni.posledni_nok_balik := "DB_HMI_recype".fronta[1].balik_den;
                   END_IF;
               END_IF;

               "DB_HMI_recype".fronta[1].prenaseny_text := '';
               "DB_HMI_recype".fronta[1].balik_den := 0;
               "DB_HMI_recype".fronta[1].vyrazeni := FALSE;

               IF #Vyrazeni.vyradit THEN
                   IF #Vyrazeni.vyrazovac_pripojen AND "DB_HMI_recype".recipe.vyrazovac_on_off THEN
                       #Vyrazeni.aktivni := TRUE;
                   ELSE
                       #Vyrazeni.alarm_nok_balik := TRUE;
                   END_IF;
               END_IF;
           END_IF;
       END_REGION

       REGION Pulz na vyrazovac - pevna delka Vyr.max_puls (200 ms)
           #TIMER.TIMER_7.TON(IN := #Vyrazeni.aktivni,
                              PT := #Vyrazeni.max_puls);
           IF #TIMER.TIMER_7.Q THEN
               #Vyrazeni.aktivni := FALSE;
           END_IF;
       END_REGION
   END_IF;

   // vystup na vyrazovac + rucni test (DB_Manual.test_vyr drzi vystup, dokud je TRUE)
   "RESERVE_DQ_2" := (#Vyrazeni.aktivni AND #Vyrazeni.vyrazovac_pripojen) OR "DB_Manual".test_vyr;

   // majak: po kazdem vyrazeni blika 5 s
   #Vyrazeni.majak_tp(IN := #Vyrazeni.aktivni AND #Vyrazeni.vyrazovac_pripojen,
                      PT := T#3S);
   #Vyrazeni.majak := #Vyrazeni.majak_tp.Q;
END_REGION

REGION Network 19 (SCL): CONTROL BLOCK presun_fronty
   IF "AUTOMAT" = true THEN


       REGION fronta 1 z 2
           IF "DB_HMI_recype".fronta[1].prenaseny_text = '' AND "DB_HMI_recype".fronta[2].prenaseny_text <> '' THEN
               "DB_HMI_recype".fronta[1]:= "DB_HMI_recype".fronta[2];
               "DB_HMI_recype".fronta[2].prenaseny_text := '';
               "DB_HMI_recype".fronta[2].balik_den := 0;
               "DB_HMI_recype".fronta[2].vyrazeni := false;
           END_IF;
       END_REGION

       REGION fronta 2 z 3
           IF "DB_HMI_recype".fronta[2].prenaseny_text = '' AND "DB_HMI_recype".fronta[3].prenaseny_text <> '' THEN
               "DB_HMI_recype".fronta[2] := "DB_HMI_recype".fronta[3];
               "DB_HMI_recype".fronta[3].prenaseny_text := '';
               "DB_HMI_recype".fronta[3].balik_den := 0;
               "DB_HMI_recype".fronta[3].vyrazeni := false;
           END_IF;
       END_REGION

       REGION fronta 3 z 4
           IF "DB_HMI_recype".fronta[3].prenaseny_text = '' AND "DB_HMI_recype".fronta[4].prenaseny_text <> '' THEN
               "DB_HMI_recype".fronta[3] := "DB_HMI_recype".fronta[4];
               "DB_HMI_recype".fronta[4].prenaseny_text := '';
               "DB_HMI_recype".fronta[4].balik_den := 0;
               "DB_HMI_recype".fronta[4].vyrazeni := false;
           END_IF;
       END_REGION

       REGION fronta 4 z 5
           IF "DB_HMI_recype".fronta[4].prenaseny_text = '' AND "DB_HMI_recype".fronta[5].prenaseny_text <> '' THEN
               "DB_HMI_recype".fronta[4] := "DB_HMI_recype".fronta[5];
               "DB_HMI_recype".fronta[5].prenaseny_text := '';
               "DB_HMI_recype".fronta[5].balik_den := 0;
               "DB_HMI_recype".fronta[5].vyrazeni := false;
           END_IF;
       END_REGION



   END_IF;


   REGION mazání fronty operátorem - bude pak možnost i automaticky ?
   IF #HMI.reset_fronty = true THEN

       "DB_HMI_recype".fronta[1].prenaseny_text := '';
       "DB_HMI_recype".fronta[1].balik_den := 0;
       "DB_HMI_recype".fronta[1].vyrazeni := false;

       "DB_HMI_recype".fronta[2].prenaseny_text := '';
       "DB_HMI_recype".fronta[2].balik_den := 0;
       "DB_HMI_recype".fronta[2].vyrazeni := false;

       "DB_HMI_recype".fronta[3].prenaseny_text := '';
       "DB_HMI_recype".fronta[3].balik_den := 0;
       "DB_HMI_recype".fronta[3].vyrazeni := false;

       "DB_HMI_recype".fronta[4].prenaseny_text := '';
       "DB_HMI_recype".fronta[4].balik_den := 0;
       "DB_HMI_recype".fronta[4].vyrazeni := false;

       "DB_HMI_recype".fronta[5].prenaseny_text := '';
       "DB_HMI_recype".fronta[5].balik_den := 0;
       "DB_HMI_recype".fronta[5].vyrazeni := false;

       "DB_HMI_recype".obsazenost_fronty := 0;
       #HMI.reset_fronty := false;

   END_IF;
   END_REGION;
END_REGION

REGION Network 20 (SCL)
   // ===== DENNI RESET POCITADLA PLAT (o pulnoci, lokalni cas) =====
   #ret := RD_LOC_T(#cas);
   IF #cas.HOUR = 0 AND #cas.MINUTE = 0 AND #cas.SECOND = 0 THEN
       #zpracovani_dat[1].balik_den := 0;
   END_IF;
   #aktual_kusy := #zpracovani_dat[1].balik_den;
END_REGION

REGION Network 21 (SCL): SBĚR VÝSLEDKŮ A ZÁPIS DO FRONTY
   #Kamera.s2_nabeh := #SENSORS.kontrola AND NOT #Kamera.s2_pamet;
   #Kamera.s2_pamet := #SENSORS.kontrola;

   IF NOT "AUTOMAT" THEN
       #Kamera.sber_aktivni := FALSE;
       #Kamera.last_id_etiketa := "COG_ETIKETA_is3800-InspectionID";
       #Kamera.last_id_folie_l := "COG_FOLIE_L_is3800-InspectionID";
       #Kamera.last_id_folie_p := "COG_FOLIE_P_is3800-InspectionID";
       #TIMER.TIMER_6.TON(IN := FALSE,
                          PT := #Kamera.timeout_sberu);
   ELSE
       REGION Prijem vysledku (zmena InspectionID = dokoncena inspekce)
           IF "COG_ETIKETA_is3800-InspectionID" <> #Kamera.last_id_etiketa THEN
               #Kamera.last_id_etiketa := "COG_ETIKETA_is3800-InspectionID";
               IF #Kamera.sber_aktivni THEN
                   #Kamera.prijato_etiketa := TRUE;
               END_IF;
           END_IF;
           // text prevzit, jakmile je k dispozici (i o par cyklu pozdeji nez ID);
           // prazdny vysledek dalsi inspekce dobry text neprepise
           IF #Kamera.sber_aktivni AND #Kamera.prijato_etiketa AND "DB_data_ctena".upraveny <> '' THEN
               #Kamera.text_etiketa := "DB_data_ctena".upraveny;
               #Kamera.ok_etiketa := TRUE;
           END_IF;
           IF "COG_FOLIE_L_is3800-InspectionID" <> #Kamera.last_id_folie_l THEN
               #Kamera.last_id_folie_l := "COG_FOLIE_L_is3800-InspectionID";
               IF #Kamera.sber_aktivni THEN
                   #Kamera.prijato_folie_l := TRUE;
                   #Kamera.ok_folie_l := ("COG_FOLIE_L_is3800-InspectionResults[0]" OR "COG_FOLIE_L_is3800-InspectionResults[1]") <> 16#00;
               END_IF;
           END_IF;
           IF "COG_FOLIE_P_is3800-InspectionID" <> #Kamera.last_id_folie_p THEN
               #Kamera.last_id_folie_p := "COG_FOLIE_P_is3800-InspectionID";
               IF #Kamera.sber_aktivni THEN
                   #Kamera.prijato_folie_p := TRUE;
                   #Kamera.ok_folie_p := ("COG_FOLIE_P_is3800-InspectionResults[0]" OR "COG_FOLIE_P_is3800-InspectionResults[1]") <> 16#00;
               END_IF;
           END_IF;
       END_REGION

       REGION Timeout - plato opustilo s2 a vysledky nedorazily
           #TIMER.TIMER_6.TON(IN := #Kamera.sber_aktivni AND NOT #SENSORS.kontrola,
                              PT := #Kamera.timeout_sberu);
       END_REGION

       REGION Vyhodnoceni a zapis do fronty
           IF #Kamera.sber_aktivni AND
               ((#Kamera.prijato_etiketa AND #Kamera.prijato_folie_l AND #Kamera.prijato_folie_p)
               OR #TIMER.TIMER_6.Q OR #Kamera.s2_nabeh) THEN

               #ocekavany_text := CONCAT(IN1 := "DB_HMI_recype".recipe.pole_string_2,
                                         IN2 := "DB_HMI_recype".recipe.pole_string_1);
               #format_etiketa_ok := #Kamera.bypass_ocr
               OR (FIND(IN1 := #Kamera.text_etiketa, IN2 := "DB_HMI_recype".recipe.pole_string_2) > 0
               AND NOT "OP2_DB".Tisk.datum_chyba);

               // kontrola kodu tridirny - nezavisla na bypass_ocr, vypinatelna z HMI
               #Kamera.tridirna_ok := NOT #Kamera.kontrola_tridirny
               OR FIND(IN1 := #Kamera.text_etiketa, IN2 := #KOD_TRIDIRNY) > 0;

               #Kamera.vyradit := NOT #Kamera.prijato_etiketa OR NOT #Kamera.prijato_folie_l
               OR NOT #Kamera.prijato_folie_p OR NOT #Kamera.ok_etiketa
               OR NOT #format_etiketa_ok OR NOT #Kamera.ok_folie_l
               OR NOT #Kamera.ok_folie_p
               OR NOT #Kamera.tridirna_ok;

               IF #Kamera.text_etiketa = '' THEN
                   #Kamera.text_etiketa := 'NECTENO';   // prazdny text = prazdna pozice!
               END_IF;

               // zapis ZA posledni obsazenou pozici
               #Kamera.idx := 0;
               FOR #i := 5 TO 1 BY -1 DO
                   IF "DB_HMI_recype".fronta[#i].prenaseny_text <> '' THEN
                       #Kamera.idx := #i;
                       EXIT;
                   END_IF;
               END_FOR;

               IF #Kamera.idx < 5 THEN
                   "DB_HMI_recype".fronta[#Kamera.idx + 1].prenaseny_text := #Kamera.text_etiketa;
                   "DB_HMI_recype".fronta[#Kamera.idx + 1].balik_den := #Kamera.balik_den;
                   "DB_HMI_recype".fronta[#Kamera.idx + 1].vyrazeni := #Kamera.vyradit;
               ELSE
                   #Kamera.fronta_plna := TRUE;
               END_IF;
               #Kamera.sber_aktivni := FALSE;
           END_IF;
       END_REGION

       REGION Novy balik pod kamerou - start sberu (az PO zapisu predchoziho)
           IF #Kamera.s2_nabeh THEN
               // citac plat (presunuto ze site 20)
               #zpracovani_dat[1].balik_den := #zpracovani_dat[1].balik_den + 1;
               IF #zpracovani_dat[1].balik_den >= 32000 THEN
                   #zpracovani_dat[1].balik_den := 1;
               END_IF;
               #Kamera.balik_den := #zpracovani_dat[1].balik_den;   // az PO pricteni

               #Kamera.sber_aktivni := TRUE;
               #Kamera.prijato_etiketa := FALSE;
               #Kamera.prijato_folie_l := FALSE;
               #Kamera.prijato_folie_p := FALSE;
               #Kamera.ok_etiketa := FALSE;
               #Kamera.ok_folie_l := FALSE;
               #Kamera.ok_folie_p := FALSE;
               #Kamera.text_etiketa := '';
           END_IF;
       END_REGION
   END_IF;

   REGION Obsazenost fronty pro HMI (pocita se kazdy scan)
       #Kamera.pocet := 0;
       FOR #i := 1 TO 5 DO
           IF "DB_HMI_recype".fronta[#i].prenaseny_text <> '' THEN
               #Kamera.pocet := #Kamera.pocet + 1;
           END_IF;
       END_FOR;
       "DB_HMI_recype".obsazenost_fronty := #Kamera.pocet;
       IF #Kamera.pocet = 0 THEN
           #Kamera.fronta_plna := FALSE;
       END_IF;
   END_REGION
END_REGION

REGION Network 22 (SCL): PŘEPNUTÍ JOBU HORNÍ KAMERY
   // Prepnuti jobu horni kamery podle receptury.
   // Spousti se nabeznou hranou "DB_HMI_recype".ODESLI_dATA (tlacitko Odeslani dat do tiskarny)
   // - soubezne s odeslanim zpravy do tiskarny (OP2).
   // Job 0 v recepture = job neprepinat.

   #Kam_Etiketa_Job.pozadovany := "DB_HMI_recype".recipe.PRG_CAM_etiketa;

   IF "CONTROL_LINE_DB".trig.reset_error_all THEN
       #Kam_Etiketa_Job.chyba := FALSE;
   END_IF;

   CASE #Kam_Etiketa_Job.krok OF
       0:  // ---- klid: cekam na pozadavek ----
           #Kam_Etiketa_Job.aktivni := FALSE;
           "COG_ETIKETA_is3800-ExecuteCommand/JobLoad" := FALSE;
           IF "DB_HMI_recype".ODESLI_dATA AND NOT #Kam_Etiketa_Job.odesli_pamet
               AND #Kam_Etiketa_Job.pozadovany > 0
               AND "COG_ETIKETA_is3800-Online" THEN
               "COG_ETIKETA_is3800-CommandID" := INT_TO_WORD(#Kam_Etiketa_Job.pozadovany);
               #Kam_Etiketa_Job.aktivni := TRUE;
               #Kam_Etiketa_Job.chyba := FALSE;
               #Kam_Etiketa_Job.krok := 10;
           END_IF;

       10: // ---- CommandID uz je venku (predchozi cyklus) -> spustit prikaz ----
           "COG_ETIKETA_is3800-ExecuteCommand/JobLoad" := TRUE;
           #Kam_Etiketa_Job.krok := 20;

       20: // ---- cekam na vysledek ----
           IF "COG_ETIKETA_is3800-CommandCompleted" THEN
               #Kam_Etiketa_Job.krok := 30;
           ELSIF "COG_ETIKETA_is3800-CommandFailed" THEN
               #Kam_Etiketa_Job.chyba := TRUE;
               #Kam_Etiketa_Job.chyba_kod := "COG_ETIKETA_is3800-CommandResultCode";
               #Kam_Etiketa_Job.krok := 30;
           ELSIF #TIMER.TIMER_3.Q THEN
               #Kam_Etiketa_Job.chyba := TRUE;            // kamera neodpovedela
               #Kam_Etiketa_Job.chyba_kod := 16#FFFF;
               #Kam_Etiketa_Job.krok := 30;
           END_IF;

